(* IEC 61131-3 sources: rusty/libs/stdlib/iec61131-st (part 2) *)

(* ---- num_conversion.st ---- *)
(********************
*
* Converts LREAL to REAL
*
*********************)
FUNCTION LREAL_TO_REAL : REAL
VAR_INPUT
    in : LREAL;
END_VAR
    LREAL_TO_REAL := in;
END_FUNCTION

(********************
*
* Converts LREAL to LINT
*
*********************)
{external}
FUNCTION LREAL_TO_LINT : LINT
VAR_INPUT
    in : LREAL;
END_VAR
END_FUNCTION

(********************
*
* Converts LREAL to DINT
*
*********************)
{external}
FUNCTION LREAL_TO_DINT : DINT
VAR_INPUT
    in : LREAL;
END_VAR
END_FUNCTION

(********************
*
* Converts LREAL to INT
*
*********************)
{external}
FUNCTION LREAL_TO_INT : INT
VAR_INPUT
    in : LREAL;
END_VAR
END_FUNCTION

(********************
*
* Converts LREAL to SINT
*
*********************)
{external}
FUNCTION LREAL_TO_SINT : SINT
VAR_INPUT
    in : LREAL;
END_VAR
END_FUNCTION

(********************
*
* Converts LREAL to ULINT
*
*********************)
{external}
FUNCTION LREAL_TO_ULINT : ULINT
VAR_INPUT
    in : LREAL;
END_VAR
END_FUNCTION

(********************
*
* Converts LREAL to UDINT
*
*********************)
{external}
FUNCTION LREAL_TO_UDINT : UDINT
VAR_INPUT
    in : LREAL;
END_VAR
END_FUNCTION

(********************
*
* Converts LREAL to UINT
*
*********************)
{external}
FUNCTION LREAL_TO_UINT : UINT
VAR_INPUT
    in : LREAL;
END_VAR
END_FUNCTION

(********************
*
* Converts LREAL to USINT
*
*********************)
{external}
FUNCTION LREAL_TO_USINT : USINT
VAR_INPUT
    in : LREAL;
END_VAR
END_FUNCTION

(********************
*
* Converts REAL to LREAL
*
*********************)
FUNCTION REAL_TO_LREAL : LREAL
VAR_INPUT
    in : REAL;
END_VAR
    REAL_TO_LREAL := in;
END_FUNCTION

(********************
*
* Converts REAL to LINT
*
*********************)
{external}
FUNCTION REAL_TO_LINT : LINT
VAR_INPUT
    in : REAL;
END_VAR
END_FUNCTION

(********************
*
* Converts REAL to DINT
*
*********************)
{external}
FUNCTION REAL_TO_DINT : DINT
VAR_INPUT
    in : REAL;
END_VAR
END_FUNCTION

(********************
*
* Converts REAL to INT
*
*********************)
{external}
FUNCTION REAL_TO_INT : INT
VAR_INPUT
    in : REAL;
END_VAR
END_FUNCTION

(********************
*
* Converts REAL to SINT
*
*********************)
{external}
FUNCTION REAL_TO_SINT : SINT
VAR_INPUT
    in : REAL;
END_VAR
END_FUNCTION

(********************
*
* Converts REAL to ULINT
*
*********************)
{external}
FUNCTION REAL_TO_ULINT : ULINT
VAR_INPUT
    in : REAL;
END_VAR
END_FUNCTION

(********************
*
* Converts REAL to UDINT
*
*********************)
{external}
FUNCTION REAL_TO_UDINT : UDINT
VAR_INPUT
    in : REAL;
END_VAR
END_FUNCTION

(********************
*
* Converts REAL to UINT
*
*********************)
{external}
FUNCTION REAL_TO_UINT : UINT
VAR_INPUT
    in : REAL;
END_VAR
END_FUNCTION

(********************
*
* Converts REAL to USINT
*
*********************)
{external}
FUNCTION REAL_TO_USINT : USINT
VAR_INPUT
    in : REAL;
END_VAR
END_FUNCTION

(********************
*
* Converts LINT to LREAL
*
*********************)
FUNCTION LINT_TO_LREAL : LREAL
VAR_INPUT
    in : LINT;
END_VAR
    LINT_TO_LREAL := in;
END_FUNCTION

(********************
*
* Converts LINT to REAL
*
*********************)
FUNCTION LINT_TO_REAL : REAL
VAR_INPUT
    in : LINT;
END_VAR
    LINT_TO_REAL := in;
END_FUNCTION

(********************
*
* Converts LINT to DINT
*
*********************)
FUNCTION LINT_TO_DINT : DINT
VAR_INPUT
    in : LINT;
END_VAR
    LINT_TO_DINT := in;
END_FUNCTION

(********************
*
* Converts LINT to INT
*
*********************)
FUNCTION LINT_TO_INT : INT
VAR_INPUT
    in : LINT;
END_VAR
    LINT_TO_INT := in;
END_FUNCTION

(********************
*
* Converts LINT to SINT
*
*********************)
FUNCTION LINT_TO_SINT : SINT
VAR_INPUT
    in : LINT;
END_VAR
    LINT_TO_SINT := in;
END_FUNCTION

(********************
*
* Converts LINT to ULINT
*
*********************)
FUNCTION LINT_TO_ULINT : ULINT
VAR_INPUT
    in : LINT;
END_VAR
    LINT_TO_ULINT := in;
END_FUNCTION

(********************
*
* Converts LINT to UDINT
*
*********************)
FUNCTION LINT_TO_UDINT : UDINT
VAR_INPUT
    in : LINT;
END_VAR
    LINT_TO_UDINT := in;
END_FUNCTION

(********************
*
* Converts LINT to UINT
*
*********************)
FUNCTION LINT_TO_UINT : UINT
VAR_INPUT
    in : LINT;
END_VAR
    LINT_TO_UINT := in;
END_FUNCTION

(********************
*
* Converts LINT to USINT
*
*********************)
FUNCTION LINT_TO_USINT : USINT
VAR_INPUT
    in : LINT;
END_VAR
    LINT_TO_USINT := in;
END_FUNCTION

(********************
*
* Converts DINT to LREAL
*
*********************)
FUNCTION DINT_TO_LREAL : LREAL
VAR_INPUT
    in : DINT;
END_VAR
    DINT_TO_LREAL := in;
END_FUNCTION

(********************
*
* Converts DINT to REAL
*
*********************)
FUNCTION DINT_TO_REAL : REAL
VAR_INPUT
    in : DINT;
END_VAR
    DINT_TO_REAL := in;
END_FUNCTION

(********************
*
* Converts DINT to LINT
*
*********************)
FUNCTION DINT_TO_LINT : LINT
VAR_INPUT
    in : DINT;
END_VAR
    DINT_TO_LINT := in;
END_FUNCTION

(********************
*
* Converts DINT to INT
*
*********************)
FUNCTION DINT_TO_INT : INT
VAR_INPUT
    in : DINT;
END_VAR
    DINT_TO_INT := in;
END_FUNCTION

(********************
*
* Converts DINT to SINT
*
*********************)
FUNCTION DINT_TO_SINT : SINT
VAR_INPUT
    in : DINT;
END_VAR
    DINT_TO_SINT := in;
END_FUNCTION

(********************
*
* Converts DINT to ULINT
*
*********************)
FUNCTION DINT_TO_ULINT : ULINT
VAR_INPUT
    in : DINT;
END_VAR
    DINT_TO_ULINT := in;
END_FUNCTION

(********************
*
* Converts DINT to UDINT
*
*********************)
FUNCTION DINT_TO_UDINT : UDINT
VAR_INPUT
    in : DINT;
END_VAR
    DINT_TO_UDINT := in;
END_FUNCTION

(********************
*
* Converts DINT to UINT
*
*********************)
FUNCTION DINT_TO_UINT : UINT
VAR_INPUT
    in : DINT;
END_VAR
    DINT_TO_UINT := in;
END_FUNCTION

(********************
*
* Converts DINT to USINT
*
*********************)
FUNCTION DINT_TO_USINT : USINT
VAR_INPUT
    in : DINT;
END_VAR
    DINT_TO_USINT := in;
END_FUNCTION

(********************
*
* Converts INT to LREAL
*
*********************)
FUNCTION INT_TO_LREAL : LREAL
VAR_INPUT
    in : INT;
END_VAR
    INT_TO_LREAL := in;
END_FUNCTION

(********************
*
* Converts INT to REAL
*
*********************)
FUNCTION INT_TO_REAL : REAL
VAR_INPUT
    in : INT;
END_VAR
    INT_TO_REAL := in;
END_FUNCTION

(********************
*
* Converts INT to LINT
*
*********************)
FUNCTION INT_TO_LINT : LINT
VAR_INPUT
    in : INT;
END_VAR
    INT_TO_LINT := in;
END_FUNCTION

(********************
*
* Converts INT to DINT
*
*********************)
FUNCTION INT_TO_DINT : DINT
VAR_INPUT
    in : INT;
END_VAR
    INT_TO_DINT := in;
END_FUNCTION

(********************
*
* Converts INT to SINT
*
*********************)
FUNCTION INT_TO_SINT : SINT
VAR_INPUT
    in : INT;
END_VAR
    INT_TO_SINT := in;
END_FUNCTION

(********************
*
* Converts INT to ULINT
*
*********************)
FUNCTION INT_TO_ULINT : ULINT
VAR_INPUT
    in : INT;
END_VAR
    INT_TO_ULINT := in;
END_FUNCTION

(********************
*
* Converts INT to UDINT
*
*********************)
FUNCTION INT_TO_UDINT : UDINT
VAR_INPUT
    in : INT;
END_VAR
    INT_TO_UDINT := in;
END_FUNCTION

(********************
*
* Converts INT to UINT
*
*********************)
FUNCTION INT_TO_UINT : UINT
VAR_INPUT
    in : INT;
END_VAR
    INT_TO_UINT := in;
END_FUNCTION

(********************
*
* Converts INT to USINT
*
*********************)
FUNCTION INT_TO_USINT : USINT
VAR_INPUT
    in : INT;
END_VAR
    INT_TO_USINT := in;
END_FUNCTION

(********************
*
* Converts SINT to LREAL
*
*********************)
FUNCTION SINT_TO_LREAL : LREAL
VAR_INPUT
    in : SINT;
END_VAR
    SINT_TO_LREAL := in;
END_FUNCTION

(********************
*
* Converts SINT to REAL
*
*********************)
FUNCTION SINT_TO_REAL : REAL
VAR_INPUT
    in : SINT;
END_VAR
    SINT_TO_REAL := in;
END_FUNCTION

(********************
*
* Converts SINT to LINT
*
*********************)
FUNCTION SINT_TO_LINT : LINT
VAR_INPUT
    in : SINT;
END_VAR
    SINT_TO_LINT := in;
END_FUNCTION

(********************
*
* Converts SINT to DINT
*
*********************)
FUNCTION SINT_TO_DINT : DINT
VAR_INPUT
    in : SINT;
END_VAR
    SINT_TO_DINT := in;
END_FUNCTION

(********************
*
* Converts SINT to INT
*
*********************)
FUNCTION SINT_TO_INT : INT
VAR_INPUT
    in : SINT;
END_VAR
    SINT_TO_INT := in;
END_FUNCTION

(********************
*
* Converts SINT to ULINT
*
*********************)
FUNCTION SINT_TO_ULINT : ULINT
VAR_INPUT
    in : SINT;
END_VAR
    SINT_TO_ULINT := in;
END_FUNCTION

(********************
*
* Converts SINT to UDINT
*
*********************)
FUNCTION SINT_TO_UDINT : UDINT
VAR_INPUT
    in : SINT;
END_VAR
    SINT_TO_UDINT := in;
END_FUNCTION

(********************
*
* Converts SINT to UINT
*
*********************)
FUNCTION SINT_TO_UINT : UINT
VAR_INPUT
    in : SINT;
END_VAR
    SINT_TO_UINT := in;
END_FUNCTION

(********************
*
* Converts SINT to USINT
*
*********************)
FUNCTION SINT_TO_USINT : USINT
VAR_INPUT
    in : SINT;
END_VAR
    SINT_TO_USINT := in;
END_FUNCTION

(********************
*
* Converts ULINT to LREAL
*
*********************)
FUNCTION ULINT_TO_LREAL : LREAL
VAR_INPUT
    in : ULINT;
END_VAR
    ULINT_TO_LREAL := in;
END_FUNCTION

(********************
*
* Converts ULINT to REAL
*
*********************)
FUNCTION ULINT_TO_REAL : REAL
VAR_INPUT
    in : ULINT;
END_VAR
    ULINT_TO_REAL := in;
END_FUNCTION

(********************
*
* Converts ULINT to LINT
*
*********************)
FUNCTION ULINT_TO_LINT : LINT
VAR_INPUT
    in : ULINT;
END_VAR
    ULINT_TO_LINT := in;
END_FUNCTION

(********************
*
* Converts ULINT to DINT
*
*********************)
FUNCTION ULINT_TO_DINT : DINT
VAR_INPUT
    in : ULINT;
END_VAR
    ULINT_TO_DINT := in;
END_FUNCTION

(********************
*
* Converts ULINT to INT
*
*********************)
FUNCTION ULINT_TO_INT : INT
VAR_INPUT
    in : ULINT;
END_VAR
    ULINT_TO_INT := in;
END_FUNCTION

(********************
*
* Converts ULINT to SINT
*
*********************)
FUNCTION ULINT_TO_SINT : SINT
VAR_INPUT
    in : ULINT;
END_VAR
    ULINT_TO_SINT := in;
END_FUNCTION

(********************
*
* Converts ULINT to UDINT
*
*********************)
FUNCTION ULINT_TO_UDINT : UDINT
VAR_INPUT
    in : ULINT;
END_VAR
    ULINT_TO_UDINT := in;
END_FUNCTION

(********************
*
* Converts ULINT to UINT
*
*********************)
FUNCTION ULINT_TO_UINT : UINT
VAR_INPUT
    in : ULINT;
END_VAR
    ULINT_TO_UINT := in;
END_FUNCTION

(********************
*
* Converts ULINT to USINT
*
*********************)
FUNCTION ULINT_TO_USINT : USINT
VAR_INPUT
    in : ULINT;
END_VAR
    ULINT_TO_USINT := in;
END_FUNCTION

(********************
*
* Converts UDINT to LREAL
*
*********************)
FUNCTION UDINT_TO_LREAL : LREAL
VAR_INPUT
    in : UDINT;
END_VAR
    UDINT_TO_LREAL := in;
END_FUNCTION

(********************
*
* Converts UDINT to REAL
*
*********************)
FUNCTION UDINT_TO_REAL : REAL
VAR_INPUT
    in : UDINT;
END_VAR
    UDINT_TO_REAL := in;
END_FUNCTION

(********************
*
* Converts UDINT to LINT
*
*********************)
FUNCTION UDINT_TO_LINT : LINT
VAR_INPUT
    in : UDINT;
END_VAR
    UDINT_TO_LINT := in;
END_FUNCTION

(********************
*
* Converts UDINT to DINT
*
*********************)
FUNCTION UDINT_TO_DINT : DINT
VAR_INPUT
    in : UDINT;
END_VAR
    UDINT_TO_DINT := in;
END_FUNCTION

(********************
*
* Converts UDINT to INT
*
*********************)
FUNCTION UDINT_TO_INT : INT
VAR_INPUT
    in : UDINT;
END_VAR
    UDINT_TO_INT := in;
END_FUNCTION

(********************
*
* Converts UDINT to SINT
*
*********************)
FUNCTION UDINT_TO_SINT : SINT
VAR_INPUT
    in : UDINT;
END_VAR
    UDINT_TO_SINT := in;
END_FUNCTION

(********************
*
* Converts UDINT to ULINT
*
*********************)
FUNCTION UDINT_TO_ULINT : ULINT
VAR_INPUT
    in : UDINT;
END_VAR
    UDINT_TO_ULINT := in;
END_FUNCTION

(********************
*
* Converts UDINT to UINT
*
*********************)
FUNCTION UDINT_TO_UINT : UINT
VAR_INPUT
    in : UDINT;
END_VAR
    UDINT_TO_UINT := in;
END_FUNCTION

(********************
*
* Converts UDINT to USINT
*
*********************)
FUNCTION UDINT_TO_USINT : USINT
VAR_INPUT
    in : UDINT;
END_VAR
    UDINT_TO_USINT := in;
END_FUNCTION

(********************
*
* Converts UINT to LREAL
*
*********************)
FUNCTION UINT_TO_LREAL : LREAL
VAR_INPUT
    in : UINT;
END_VAR
    UINT_TO_LREAL := in;
END_FUNCTION

(********************
*
* Converts UINT to REAL
*
*********************)
FUNCTION UINT_TO_REAL : REAL
VAR_INPUT
    in : UINT;
END_VAR
    UINT_TO_REAL := in;
END_FUNCTION

(********************
*
* Converts UINT to LINT
*
*********************)
FUNCTION UINT_TO_LINT : LINT
VAR_INPUT
    in : UINT;
END_VAR
    UINT_TO_LINT := in;
END_FUNCTION

(********************
*
* Converts UINT to DINT
*
*********************)
FUNCTION UINT_TO_DINT : DINT
VAR_INPUT
    in : UINT;
END_VAR
    UINT_TO_DINT := in;
END_FUNCTION

(********************
*
* Converts UINT to INT
*
*********************)
FUNCTION UINT_TO_INT : INT
VAR_INPUT
    in : UINT;
END_VAR
    UINT_TO_INT := in;
END_FUNCTION

(********************
*
* Converts UINT to SINT
*
*********************)
FUNCTION UINT_TO_SINT : SINT
VAR_INPUT
    in : UINT;
END_VAR
    UINT_TO_SINT := in;
END_FUNCTION

(********************
*
* Converts UINT to ULINT
*
*********************)
FUNCTION UINT_TO_ULINT : ULINT
VAR_INPUT
    in : UINT;
END_VAR
    UINT_TO_ULINT := in;
END_FUNCTION

(********************
*
* Converts UINT to UDINT
*
*********************)
FUNCTION UINT_TO_UDINT : UDINT
VAR_INPUT
    in : UINT;
END_VAR
    UINT_TO_UDINT := in;
END_FUNCTION

(********************
*
* Converts UINT to USINT
*
*********************)
FUNCTION UINT_TO_USINT : USINT
VAR_INPUT
    in : UINT;
END_VAR
    UINT_TO_USINT := in;
END_FUNCTION

(********************
*
* Converts USINT to LREAL
*
*********************)
FUNCTION USINT_TO_LREAL : LREAL
VAR_INPUT
    in : USINT;
END_VAR
    USINT_TO_LREAL := in;
END_FUNCTION

(********************
*
* Converts USINT to REAL
*
*********************)
FUNCTION USINT_TO_REAL : REAL
VAR_INPUT
    in : USINT;
END_VAR
    USINT_TO_REAL := in;
END_FUNCTION

(********************
*
* Converts USINT to LINT
*
*********************)
FUNCTION USINT_TO_LINT : LINT
VAR_INPUT
    in : USINT;
END_VAR
    USINT_TO_LINT := in;
END_FUNCTION

(********************
*
* Converts USINT to DINT
*
*********************)
FUNCTION USINT_TO_DINT : DINT
VAR_INPUT
    in : USINT;
END_VAR
    USINT_TO_DINT := in;
END_FUNCTION

(********************
*
* Converts USINT to INT
*
*********************)
FUNCTION USINT_TO_INT : INT
VAR_INPUT
    in : USINT;
END_VAR
    USINT_TO_INT := in;
END_FUNCTION

(********************
*
* Converts USINT to SINT
*
*********************)
FUNCTION USINT_TO_SINT : SINT
VAR_INPUT
    in : USINT;
END_VAR
    USINT_TO_SINT := in;
END_FUNCTION

(********************
*
* Converts USINT to ULINT
*
*********************)
FUNCTION USINT_TO_ULINT : ULINT
VAR_INPUT
    in : USINT;
END_VAR
    USINT_TO_ULINT := in;
END_FUNCTION

(********************
*
* Converts USINT to UDINT
*
*********************)
FUNCTION USINT_TO_UDINT : UDINT
VAR_INPUT
    in : USINT;
END_VAR
    USINT_TO_UDINT := in;
END_FUNCTION

(********************
*
* Converts USINT to UINT
*
*********************)
FUNCTION USINT_TO_UINT : UINT
VAR_INPUT
    in : USINT;
END_VAR
    USINT_TO_UINT := in;
END_FUNCTION

(* ---- numerical_functions.st ---- *)
(**************************
 *
 *This operator returns the absolute value of a number.
 *
*************************)
FUNCTION ABS<T : ANY_NUM> : T
VAR_INPUT
    IN : T;
END_VAR

END_FUNCTION

(* Specialized implementation of ABS for DINT *)
/* FUNCTION ABS__DINT : DINT */
FUNCTION ABS__DINT : DINT
VAR_INPUT
    IN : DINT;
END_VAR
    ABS__DINT := IN;
    IF ABS__DINT < 0 THEN
        ABS__DINT := -1 * ABS__DINT;
    END_IF
END_FUNCTION

(* Specialized implementation of ABS for SINT *)
FUNCTION ABS__SINT : SINT
VAR_INPUT
    IN : SINT;
END_VAR
    ABS__SINT := ABS__DINT(IN);
END_FUNCTION

(* Specialized implementation of ABS for INT *)
FUNCTION ABS__INT : INT
VAR_INPUT
    IN : INT;
END_VAR
    ABS__INT := ABS__DINT(IN);
END_FUNCTION

(* Specialized implementation of ABS for LINT *)
FUNCTION ABS__LINT : LINT
VAR_INPUT
    IN : LINT;
END_VAR
    ABS__LINT := IN;
    IF ABS__LINT < 0 THEN
        ABS__LINT := -1 * ABS__LINT;
    END_IF
END_FUNCTION

(* Specialized implementation of ABS for REAL *)
FUNCTION ABS__REAL : REAL
VAR_INPUT
    IN : REAL;
END_VAR
    ABS__REAL := ABS__LREAL(IN);
END_FUNCTION

(* Specialized implementation of ABS for LREAL *)
FUNCTION ABS__LREAL : LREAL
VAR_INPUT
    IN : LREAL;
END_VAR
    ABS__LREAL := IN;
    IF ABS__LREAL < 0 THEN
        ABS__LREAL := -1.0 * ABS__LREAL;
    END_IF
END_FUNCTION

(* ---- real_trunc_int.st ---- *)
(********************
*
* Converts REAL to SINT
*
********************)
FUNCTION REAL_TRUNC_SINT : SINT
    VAR_INPUT
        in : REAL;
    END_VAR

    REAL_TRUNC_SINT := in;
END_FUNCTION

(********************
*
* Converts REAL to USINT
*
********************)
FUNCTION REAL_TRUNC_USINT : USINT
    VAR_INPUT
        in : REAL;
    END_VAR

    REAL_TRUNC_USINT := in;
END_FUNCTION

(********************
*
* Converts REAL to INT
*
********************)
FUNCTION REAL_TRUNC_INT : INT
    VAR_INPUT
        in : REAL;
    END_VAR

    REAL_TRUNC_INT := in;
END_FUNCTION

(********************
*
* Converts REAL to UINT
*
********************)
FUNCTION REAL_TRUNC_UINT : UINT
    VAR_INPUT
        in : REAL;
    END_VAR

    REAL_TRUNC_UINT := in;
END_FUNCTION

(********************
*
* Converts REAL to DINT
*
********************)
FUNCTION REAL_TRUNC_DINT : DINT
    VAR_INPUT
        in : REAL;
    END_VAR

    REAL_TRUNC_DINT := in;
END_FUNCTION

(********************
*
* Converts REAL to UDINT
*
********************)
FUNCTION REAL_TRUNC_UDINT : UDINT
    VAR_INPUT
        in : REAL;
    END_VAR

    REAL_TRUNC_UDINT := in;
END_FUNCTION

(********************
*
* Converts REAL to LINT
*
********************)
FUNCTION REAL_TRUNC_LINT : LINT
    VAR_INPUT
        in : REAL;
    END_VAR

    REAL_TRUNC_LINT := in;
END_FUNCTION

(********************
*
* Converts REAL to ULINT
*
********************)
FUNCTION REAL_TRUNC_ULINT : ULINT
    VAR_INPUT
        in : REAL;
    END_VAR

    REAL_TRUNC_ULINT := in;
END_FUNCTION

(********************
*
* Converts LREAL to SINT
*
********************)
FUNCTION LREAL_TRUNC_SINT : SINT
    VAR_INPUT
        in : LREAL;
    END_VAR

    LREAL_TRUNC_SINT := in;
END_FUNCTION

(********************
*
* Converts LREAL to USINT
*
********************)
FUNCTION LREAL_TRUNC_USINT : USINT
    VAR_INPUT
        in : LREAL;
    END_VAR

    LREAL_TRUNC_USINT := in;
END_FUNCTION

(********************
*
* Converts LREAL to INT
*
********************)
FUNCTION LREAL_TRUNC_INT : INT
    VAR_INPUT
        in : LREAL;
    END_VAR

    LREAL_TRUNC_INT := in;
END_FUNCTION

(********************
*
* Converts LREAL to UINT
*
********************)
FUNCTION LREAL_TRUNC_UINT : UINT
    VAR_INPUT
        in : LREAL;
    END_VAR

    LREAL_TRUNC_UINT := in;
END_FUNCTION

(********************
*
* Converts LREAL to DINT
*
********************)
FUNCTION LREAL_TRUNC_DINT : DINT
    VAR_INPUT
        in : LREAL;
    END_VAR

    LREAL_TRUNC_DINT := in;
END_FUNCTION

(********************
*
* Converts LREAL to UDINT
*
********************)
FUNCTION LREAL_TRUNC_UDINT : UDINT
    VAR_INPUT
        in : LREAL;
    END_VAR

    LREAL_TRUNC_UDINT := in;
END_FUNCTION

(********************
*
* Converts LREAL to LINT
*
********************)
FUNCTION LREAL_TRUNC_LINT : LINT
    VAR_INPUT
        in : LREAL;
    END_VAR

    LREAL_TRUNC_LINT := in;
END_FUNCTION

(********************
*
* Converts LREAL to ULINT
*
********************)
FUNCTION LREAL_TRUNC_ULINT : ULINT
    VAR_INPUT
        in : LREAL;
    END_VAR

    LREAL_TRUNC_ULINT := in;
END_FUNCTION

(* ---- selectors.st ---- *)
(**************************
 *
 * MAX(IN0, IN1, ...)
 *
 * This operator produces the larger value of the given operands.
 *
*************************)
{external}
FUNCTION MAX<T: ANY_ELEMENTARY> : T
VAR_INPUT
    IN : {sized} T...;
END_VAR
END_FUNCTION

(**************************
 *
 * MIN(IN0, IN1, ...)
 *
 * This operator produces the smaller value of the given operands.
 *
*************************)
{external}
FUNCTION MIN<T: ANY_ELEMENTARY> : T
VAR_INPUT
    IN : {sized} T...;
END_VAR
END_FUNCTION

(**************************
 *
 * LIMIT(Min, IN, Max)
 *
 * This operator limits an input value to the range between Min and Max.
 * If IN lies between the range of Min and Max, IN is displayed as a result.
 * If IN > Max, Max is displayed as a result.
 * If IN < Min, Min is displayed as a result.
 *
*************************)
{external}
FUNCTION LIMIT<T: ANY_ELEMENTARY> : T
VAR_INPUT
    MIN : T;
    IN : T;
    MAX : T;
END_VAR
END_FUNCTION

(* ---- string_conversion.st ---- *)
(********************
*
* Converts WSTRING to STRING
*
*********************)
FUNCTION WSTRING_TO_STRING : STRING[__STRING_LENGTH]
VAR_INPUT {ref}
    in : WSTRING[__STRING_LENGTH];
END_VAR
    WSTRING_TO_STRING_EXT(in, WSTRING_TO_STRING);
END_FUNCTION

{external}
FUNCTION WSTRING_TO_STRING_EXT : DINT
VAR_INPUT {ref}
    in : WSTRING[__STRING_LENGTH];
END_VAR
VAR_IN_OUT
    out : STRING[__STRING_LENGTH];
END_VAR
END_FUNCTION

(********************
*
* Converts WSTRING to WCHAR
*
*********************)
{external}
FUNCTION WSTRING_TO_WCHAR : WCHAR
VAR_INPUT {ref}
    in : WSTRING;
END_VAR
END_FUNCTION

(********************
*
* Converts STRING to WSTRING
* Will return a WSTRING with default length of 81
*
*********************)
FUNCTION STRING_TO_WSTRING : WSTRING[__STRING_LENGTH]
VAR_INPUT {ref}
    in : STRING[__STRING_LENGTH];
END_VAR
    STRING_TO_WSTRING_EXT(in, STRING_TO_WSTRING);
END_FUNCTION

{external}
FUNCTION STRING_TO_WSTRING_EXT : DINT
VAR_INPUT {ref}
    in : STRING[__STRING_LENGTH];
END_VAR
VAR_IN_OUT
    out : WSTRING[__STRING_LENGTH];
END_VAR
END_FUNCTION

(********************
*
* Converts STRING to CHAR
*
*********************)
{external}
FUNCTION STRING_TO_CHAR : CHAR
VAR_INPUT {ref}
    in : STRING;
END_VAR
END_FUNCTION

(********************
*
* Converts WCHAR to WSTRING
*
*********************)
{external}
FUNCTION WCHAR_TO_WSTRING : WSTRING
VAR_INPUT
    in : WCHAR;
END_VAR
END_FUNCTION

(********************
*
* Converts WCHAR to CHAR
*
*********************)
{external}
FUNCTION WCHAR_TO_CHAR : CHAR
VAR_INPUT
    in : WCHAR;
END_VAR
END_FUNCTION

(********************
*
* Converts CHAR to STRING
*
*********************)
{external}
FUNCTION CHAR_TO_STRING : STRING
VAR_INPUT
    in : CHAR;
END_VAR
END_FUNCTION

(********************
*
* Converts CHAR to WCHAR
*
*********************)
{external}
FUNCTION CHAR_TO_WCHAR : WCHAR
VAR_INPUT
    in : CHAR;
END_VAR
END_FUNCTION

(* ---- string_to_conversions.st ---- *)
(******************************************************************************
*
* Converts STRING and WSTRING values to native values.
*
******************************************************************************)

(******************************************************************************
*
* Converts STRING to BOOL. Never faults; a rejected input yields FALSE.
*
******************************************************************************)
{external}
FUNCTION STRING_TO_BOOL : BOOL
VAR_INPUT {ref}
    IN : STRING;
END_VAR
END_FUNCTION

(******************************************************************************
*
* Converts STRING to BYTE. Never faults; a rejected input yields 0.
*
******************************************************************************)
{external}
FUNCTION STRING_TO_BYTE : BYTE
VAR_INPUT {ref}
    IN : STRING;
END_VAR
END_FUNCTION

(******************************************************************************
*
* Converts STRING to WORD. Never faults; a rejected input yields 0.
*
******************************************************************************)
{external}
FUNCTION STRING_TO_WORD : WORD
VAR_INPUT {ref}
    IN : STRING;
END_VAR
END_FUNCTION

(******************************************************************************
*
* Converts STRING to DWORD. Never faults; a rejected input yields 0.
*
******************************************************************************)
{external}
FUNCTION STRING_TO_DWORD : DWORD
VAR_INPUT {ref}
    IN : STRING;
END_VAR
END_FUNCTION

(******************************************************************************
*
* Converts STRING to LWORD. Never faults; a rejected input yields 0.
*
******************************************************************************)
{external}
FUNCTION STRING_TO_LWORD : LWORD
VAR_INPUT {ref}
    IN : STRING;
END_VAR
END_FUNCTION

(******************************************************************************
*
* Converts STRING to SINT. Never faults; a rejected input yields 0.
*
******************************************************************************)
{external}
FUNCTION STRING_TO_SINT : SINT
VAR_INPUT {ref}
    IN : STRING;
END_VAR
END_FUNCTION

(******************************************************************************
*
* Converts STRING to USINT. Never faults; a rejected input yields 0.
*
******************************************************************************)
{external}
FUNCTION STRING_TO_USINT : USINT
VAR_INPUT {ref}
    IN : STRING;
END_VAR
END_FUNCTION

(******************************************************************************
*
* Converts STRING to INT. Never faults; a rejected input yields 0.
*
******************************************************************************)
{external}
FUNCTION STRING_TO_INT : INT
VAR_INPUT {ref}
    IN : STRING;
END_VAR
END_FUNCTION

(******************************************************************************
*
* Converts STRING to UINT. Never faults; a rejected input yields 0.
*
******************************************************************************)
{external}
FUNCTION STRING_TO_UINT : UINT
VAR_INPUT {ref}
    IN : STRING;
END_VAR
END_FUNCTION

(******************************************************************************
*
* Converts STRING to DINT. Never faults; a rejected input yields 0.
*
******************************************************************************)
{external}
FUNCTION STRING_TO_DINT : DINT
VAR_INPUT {ref}
    IN : STRING;
END_VAR
END_FUNCTION

(******************************************************************************
*
* Converts STRING to UDINT. Never faults; a rejected input yields 0.
*
******************************************************************************)
{external}
FUNCTION STRING_TO_UDINT : UDINT
VAR_INPUT {ref}
    IN : STRING;
END_VAR
END_FUNCTION

(******************************************************************************
*
* Converts STRING to LINT. Never faults; a rejected input yields 0.
*
******************************************************************************)
{external}
FUNCTION STRING_TO_LINT : LINT
VAR_INPUT {ref}
    IN : STRING;
END_VAR
END_FUNCTION

(******************************************************************************
*
* Converts STRING to ULINT. Never faults; a rejected input yields 0.
*
******************************************************************************)
{external}
FUNCTION STRING_TO_ULINT : ULINT
VAR_INPUT {ref}
    IN : STRING;
END_VAR
END_FUNCTION

(******************************************************************************
*
* Converts STRING to LREAL.
*
******************************************************************************)
{external}
FUNCTION STRING_TO_LREAL : LREAL
VAR_INPUT {ref}
    IN : STRING;
END_VAR
END_FUNCTION

(******************************************************************************
*
* Converts STRING to REAL.
*
******************************************************************************)
{external}
FUNCTION STRING_TO_REAL : REAL
VAR_INPUT {ref}
    IN : STRING;
END_VAR
END_FUNCTION

(******************************************************************************
*
* Converts STRING to TIME. Requires a T#/TIME# prefix; never faults, a rejected or
* negative duration yields T#0s.
*
******************************************************************************)
{external}
FUNCTION STRING_TO_TIME : TIME
VAR_INPUT {ref}
    IN : STRING;
END_VAR
END_FUNCTION

(******************************************************************************
*
* Converts STRING to LTIME. Requires a LT#/LTIME# prefix; never faults, a rejected or
* negative duration yields LTIME#0s.
*
******************************************************************************)
{external}
FUNCTION STRING_TO_LTIME : LTIME
VAR_INPUT {ref}
    IN : STRING;
END_VAR
END_FUNCTION

(******************************************************************************
*
* Converts STRING to DATE. Requires a D#/DATE# prefix. Never faults; an impossible or
* out-of-range (1970-01-01..2106-02-07) date yields D#1970-01-01.
*
******************************************************************************)
{external}
FUNCTION STRING_TO_DATE : DATE
VAR_INPUT {ref}
    IN : STRING;
END_VAR
END_FUNCTION

(******************************************************************************
*
* Converts STRING to DT. Requires a DT#/DATE_AND_TIME# prefix. Never faults; an
* impossible or out-of-range date-time yields DT#1970-01-01-00:00:00.
*
******************************************************************************)
{external}
FUNCTION STRING_TO_DT : DT
VAR_INPUT {ref}
    IN : STRING;
END_VAR
END_FUNCTION

(******************************************************************************
*
* Converts STRING to TOD. Requires a TOD#/TIME_OF_DAY# prefix. Never faults; an
* impossible time yields TOD#00:00:00.
*
******************************************************************************)
{external}
FUNCTION STRING_TO_TOD : TOD
VAR_INPUT {ref}
    IN : STRING;
END_VAR
END_FUNCTION

(******************************************************************************
*
* Converts WSTRING to LINT.
*
******************************************************************************)
FUNCTION WSTRING_TO_LINT : LINT
VAR_INPUT {ref}
    IN : WSTRING;
END_VAR
VAR_TEMP
    STR : STRING;
END_VAR
    WSTRING_TO_STRING_EXT(IN, STR);
    WSTRING_TO_LINT := STRING_TO_LINT(STR);
END_FUNCTION

(******************************************************************************
*
* Converts WSTRING to DINT.
*
******************************************************************************)
FUNCTION WSTRING_TO_DINT : DINT
VAR_INPUT {ref}
    IN : WSTRING;
END_VAR
VAR_TEMP
    STR : STRING;
END_VAR
    WSTRING_TO_STRING_EXT(IN, STR);
    WSTRING_TO_DINT := STRING_TO_DINT(STR);
END_FUNCTION

(******************************************************************************
*
* Converts WSTRING to LREAL.
*
******************************************************************************)
FUNCTION WSTRING_TO_LREAL : LREAL
VAR_INPUT {ref}
    IN : WSTRING;
END_VAR
VAR_TEMP
    STR : STRING;
END_VAR
    WSTRING_TO_STRING_EXT(IN, STR);
    WSTRING_TO_LREAL := STRING_TO_LREAL(STR);
END_FUNCTION

(******************************************************************************
*
* Converts WSTRING to REAL.
*
******************************************************************************)
FUNCTION WSTRING_TO_REAL : REAL
VAR_INPUT {ref}
    IN : WSTRING;
END_VAR
VAR_TEMP
    STR : STRING;
END_VAR
    WSTRING_TO_STRING_EXT(IN, STR);
    WSTRING_TO_REAL := STRING_TO_REAL(STR);
END_FUNCTION

(* ---- to_bit.st ---- *)
FUNCTION TO_BOOL<T: ANY> : BOOL
    VAR_INPUT
        in : T;
    END_VAR
END_FUNCTION

FUNCTION TO_BOOL__BOOL : BOOL
    VAR_INPUT
        in : BOOL;
    END_VAR

    TO_BOOL__BOOL := in;
END_FUNCTION

FUNCTION TO_BOOL__BYTE : BOOL
    VAR_INPUT
        in : BYTE;
    END_VAR

    TO_BOOL__BYTE := BYTE_TO_BOOL(in);
END_FUNCTION

FUNCTION TO_BOOL__WORD : BOOL
    VAR_INPUT
        in : WORD;
    END_VAR

    TO_BOOL__WORD := WORD_TO_BOOL(in);
END_FUNCTION

FUNCTION TO_BOOL__DWORD : BOOL
    VAR_INPUT
        in : DWORD;
    END_VAR

    TO_BOOL__DWORD := DWORD_TO_BOOL(in);
END_FUNCTION

FUNCTION TO_BOOL__LWORD : BOOL
    VAR_INPUT
        in : LWORD;
    END_VAR

    TO_BOOL__LWORD := LWORD_TO_BOOL(in);
END_FUNCTION

FUNCTION TO_BOOL__SINT : BOOL
    VAR_INPUT
        in : SINT;
    END_VAR

    TO_BOOL__SINT := SINT_TO_BOOL(in);
END_FUNCTION

FUNCTION TO_BOOL__USINT : BOOL
    VAR_INPUT
        in : USINT;
    END_VAR

    TO_BOOL__USINT := USINT_TO_BOOL(in);
END_FUNCTION

FUNCTION TO_BOOL__INT : BOOL
    VAR_INPUT
        in : INT;
    END_VAR

    TO_BOOL__INT := INT_TO_BOOL(in);
END_FUNCTION

FUNCTION TO_BOOL__UINT : BOOL
    VAR_INPUT
        in : UINT;
    END_VAR

    TO_BOOL__UINT := UINT_TO_BOOL(in);
END_FUNCTION

FUNCTION TO_BOOL__DINT : BOOL
    VAR_INPUT
        in : DINT;
    END_VAR

    TO_BOOL__DINT := DINT_TO_BOOL(in);
END_FUNCTION

FUNCTION TO_BOOL__UDINT : BOOL
    VAR_INPUT
        in : UDINT;
    END_VAR

    TO_BOOL__UDINT := UDINT_TO_BOOL(in);
END_FUNCTION

FUNCTION TO_BOOL__LINT : BOOL
    VAR_INPUT
        in : LINT;
    END_VAR

    TO_BOOL__LINT := LINT_TO_BOOL(in);
END_FUNCTION

FUNCTION TO_BOOL__ULINT : BOOL
    VAR_INPUT
        in : ULINT;
    END_VAR

    TO_BOOL__ULINT := ULINT_TO_BOOL(in);
END_FUNCTION

FUNCTION TO_BOOL__REAL : BOOL
    VAR_INPUT
        in : REAL;
    END_VAR

    TO_BOOL__REAL := REAL_TO_BOOL(in);
END_FUNCTION

FUNCTION TO_BOOL__LREAL : BOOL
    VAR_INPUT
        in : LREAL;
    END_VAR

    TO_BOOL__LREAL := LREAL_TO_BOOL(in);
END_FUNCTION

// ======================================================================================================== //

FUNCTION TO_BYTE<T: ANY> : BYTE
    VAR_INPUT
        in : T;
    END_VAR
END_FUNCTION

FUNCTION TO_BYTE__BYTE : BYTE
    VAR_INPUT
        in : BYTE;
    END_VAR

    TO_BYTE__BYTE := in;
END_FUNCTION

FUNCTION TO_BYTE__BOOL : BYTE
    VAR_INPUT
        in : BOOL;
    END_VAR

    TO_BYTE__BOOL := BOOL_TO_BYTE(in);
END_FUNCTION

FUNCTION TO_BYTE__CHAR : BYTE
    VAR_INPUT
        in : CHAR;
    END_VAR

    TO_BYTE__CHAR := CHAR_TO_BYTE(in);
END_FUNCTION

FUNCTION TO_BYTE__WCHAR : BYTE
    VAR_INPUT
        in : WCHAR;
    END_VAR

    TO_BYTE__WCHAR := WCHAR_TO_BYTE(in);
END_FUNCTION

FUNCTION TO_BYTE__WORD : BYTE
    VAR_INPUT
        in : WORD;
    END_VAR

    TO_BYTE__WORD := WORD_TO_BYTE(in);
END_FUNCTION

FUNCTION TO_BYTE__DWORD : BYTE
    VAR_INPUT
        in : DWORD;
    END_VAR

    TO_BYTE__DWORD := DWORD_TO_BYTE(in);
END_FUNCTION

FUNCTION TO_BYTE__LWORD : BYTE
    VAR_INPUT
        in : LWORD;
    END_VAR

    TO_BYTE__LWORD := LWORD_TO_BYTE(in);
END_FUNCTION

FUNCTION TO_BYTE__REAL : BYTE
    VAR_INPUT
        in : REAL;
    END_VAR

    TO_BYTE__REAL := REAL_TO_BYTE(in);
END_FUNCTION

FUNCTION TO_BYTE__LREAL : BYTE
    VAR_INPUT
        in : LREAL;
    END_VAR

    TO_BYTE__LREAL := LREAL_TO_BYTE(in);
END_FUNCTION

// ======================================================================================================== //

FUNCTION TO_WORD<T: ANY> : WORD
    VAR_INPUT
        in : T;
    END_VAR
END_FUNCTION

FUNCTION TO_WORD__WORD : WORD
    VAR_INPUT
        in : WORD;
    END_VAR

    TO_WORD__WORD := in;
END_FUNCTION

FUNCTION TO_WORD__BOOL : WORD
    VAR_INPUT
        in : BOOL;
    END_VAR

    TO_WORD__BOOL := BOOL_TO_WORD(in);
END_FUNCTION

FUNCTION TO_WORD__CHAR : WORD
    VAR_INPUT
        in : CHAR;
    END_VAR

    TO_WORD__CHAR := CHAR_TO_WORD(in);
END_FUNCTION

FUNCTION TO_WORD__WCHAR : WORD
    VAR_INPUT
        in : WCHAR;
    END_VAR

    TO_WORD__WCHAR := WCHAR_TO_WORD(in);
END_FUNCTION

FUNCTION TO_WORD__BYTE : WORD
    VAR_INPUT
        in : BYTE;
    END_VAR

    TO_WORD__BYTE := BYTE_TO_WORD(in);
END_FUNCTION

FUNCTION TO_WORD__DWORD : WORD
    VAR_INPUT
        in : DWORD;
    END_VAR

    TO_WORD__DWORD := DWORD_TO_WORD(in);
END_FUNCTION

FUNCTION TO_WORD__LWORD : WORD
    VAR_INPUT
        in : LWORD;
    END_VAR

    TO_WORD__LWORD := LWORD_TO_WORD(in);
END_FUNCTION

FUNCTION TO_WORD__REAL : WORD
    VAR_INPUT
        in : REAL;
    END_VAR

    TO_WORD__REAL := REAL_TO_WORD(in);
END_FUNCTION

FUNCTION TO_WORD__LREAL : WORD
    VAR_INPUT
        in : LREAL;
    END_VAR

    TO_WORD__LREAL := LREAL_TO_WORD(in);
END_FUNCTION

// ======================================================================================================== //

FUNCTION TO_DWORD<T: ANY> : DWORD
    VAR_INPUT
        in : T;
    END_VAR
END_FUNCTION

FUNCTION TO_DWORD__DWORD : DWORD
    VAR_INPUT
        in : DWORD;
    END_VAR

    TO_DWORD__DWORD := in;
END_FUNCTION

FUNCTION TO_DWORD__BOOL : DWORD
    VAR_INPUT
        in : BOOL;
    END_VAR

    TO_DWORD__BOOL := BOOL_TO_DWORD(in);
END_FUNCTION

FUNCTION TO_DWORD__CHAR : DWORD
    VAR_INPUT
        in : CHAR;
    END_VAR

    TO_DWORD__CHAR := CHAR_TO_DWORD(in);
END_FUNCTION

FUNCTION TO_DWORD__WCHAR : DWORD
    VAR_INPUT
        in : WCHAR;
    END_VAR

    TO_DWORD__WCHAR := WCHAR_TO_DWORD(in);
END_FUNCTION

FUNCTION TO_DWORD__BYTE : DWORD
    VAR_INPUT
        in : BYTE;
    END_VAR

    TO_DWORD__BYTE := BYTE_TO_DWORD(in);
END_FUNCTION

FUNCTION TO_DWORD__WORD : DWORD
    VAR_INPUT
        in : WORD;
    END_VAR

    TO_DWORD__WORD := WORD_TO_DWORD(in);
END_FUNCTION

FUNCTION TO_DWORD__LWORD : DWORD
    VAR_INPUT
        in : LWORD;
    END_VAR

    TO_DWORD__LWORD := LWORD_TO_DWORD(in);
END_FUNCTION

FUNCTION TO_DWORD__REAL : DWORD
    VAR_INPUT
        in : REAL;
    END_VAR

    TO_DWORD__REAL := REAL_TO_DWORD(in);
END_FUNCTION

FUNCTION TO_DWORD__LREAL : DWORD
    VAR_INPUT
        in : LREAL;
    END_VAR

    TO_DWORD__LREAL := LREAL_TO_DWORD(in);
END_FUNCTION

// ======================================================================================================== //

FUNCTION TO_LWORD<T: ANY> : LWORD
    VAR_INPUT
        in : T;
    END_VAR
END_FUNCTION

FUNCTION TO_LWORD__LWORD : LWORD
    VAR_INPUT
        in : LWORD;
    END_VAR

    TO_LWORD__LWORD := in;
END_FUNCTION

FUNCTION TO_LWORD__BOOL : LWORD
    VAR_INPUT
        in : BOOL;
    END_VAR

    TO_LWORD__BOOL := BOOL_TO_LWORD(in);
END_FUNCTION

FUNCTION TO_LWORD__CHAR : LWORD
    VAR_INPUT
        in : CHAR;
    END_VAR

    TO_LWORD__CHAR := CHAR_TO_LWORD(in);
END_FUNCTION

FUNCTION TO_LWORD__WCHAR : LWORD
    VAR_INPUT
        in : WCHAR;
    END_VAR

    TO_LWORD__WCHAR := WCHAR_TO_LWORD(in);
END_FUNCTION

FUNCTION TO_LWORD__BYTE : LWORD
    VAR_INPUT
        in : BYTE;
    END_VAR

    TO_LWORD__BYTE := BYTE_TO_LWORD(in);
END_FUNCTION

FUNCTION TO_LWORD__WORD : LWORD
    VAR_INPUT
        in : WORD;
    END_VAR

    TO_LWORD__WORD := WORD_TO_LWORD(in);
END_FUNCTION

FUNCTION TO_LWORD__DWORD : LWORD
    VAR_INPUT
        in : DWORD;
    END_VAR

    TO_LWORD__DWORD := DWORD_TO_LWORD(in);
END_FUNCTION

FUNCTION TO_LWORD__REAL : LWORD
    VAR_INPUT
        in : REAL;
    END_VAR

    TO_LWORD__REAL := REAL_TO_LWORD(in);
END_FUNCTION

FUNCTION TO_LWORD__LREAL : LWORD
    VAR_INPUT
        in : LREAL;
    END_VAR

    TO_LWORD__LREAL := LREAL_TO_LWORD(in);
END_FUNCTION

(* ---- to_date_time.st ---- *)
FUNCTION TO_TIME<T: ANY> : TIME
    VAR_INPUT
        in : T;
    END_VAR
END_FUNCTION

FUNCTION TO_TIME__TIME : TIME
    VAR_INPUT
        in : TIME;
    END_VAR

    TO_TIME__TIME := in;
END_FUNCTION

FUNCTION TO_TIME__LTIME : TIME
    VAR_INPUT
        in : LTIME;
    END_VAR

    TO_TIME__LTIME := LTIME_TO_TIME(in);
END_FUNCTION

FUNCTION TO_TIME__BOOL : TIME
    VAR_INPUT
        in : BOOL;
    END_VAR

    TO_TIME__BOOL := BOOL_TO_TIME(in);
END_FUNCTION

FUNCTION TO_TIME__BYTE : TIME
    VAR_INPUT
        in : BYTE;
    END_VAR

    TO_TIME__BYTE := BYTE_TO_TIME(in);
END_FUNCTION

FUNCTION TO_TIME__WORD : TIME
    VAR_INPUT
        in : WORD;
    END_VAR

    TO_TIME__WORD := WORD_TO_TIME(in);
END_FUNCTION

FUNCTION TO_TIME__DWORD : TIME
    VAR_INPUT
        in : DWORD;
    END_VAR

    TO_TIME__DWORD := DWORD_TO_TIME(in);
END_FUNCTION

FUNCTION TO_TIME__LWORD : TIME
    VAR_INPUT
        in : LWORD;
    END_VAR

    TO_TIME__LWORD := LWORD_TO_TIME(in);
END_FUNCTION

FUNCTION TO_TIME__SINT : TIME
    VAR_INPUT
        in : SINT;
    END_VAR

    TO_TIME__SINT := SINT_TO_TIME(in);
END_FUNCTION

FUNCTION TO_TIME__USINT : TIME
    VAR_INPUT
        in : USINT;
    END_VAR

    TO_TIME__USINT := USINT_TO_TIME(in);
END_FUNCTION

FUNCTION TO_TIME__INT : TIME
    VAR_INPUT
        in : INT;
    END_VAR

    TO_TIME__INT := INT_TO_TIME(in);
END_FUNCTION

FUNCTION TO_TIME__UINT : TIME
    VAR_INPUT
        in : UINT;
    END_VAR

    TO_TIME__UINT := UINT_TO_TIME(in);
END_FUNCTION

FUNCTION TO_TIME__DINT : TIME
    VAR_INPUT
        in : DINT;
    END_VAR

    TO_TIME__DINT := DINT_TO_TIME(in);
END_FUNCTION

FUNCTION TO_TIME__UDINT : TIME
    VAR_INPUT
        in : UDINT;
    END_VAR

    TO_TIME__UDINT := UDINT_TO_TIME(in);
END_FUNCTION

FUNCTION TO_TIME__LINT : TIME
    VAR_INPUT
        in : LINT;
    END_VAR

    TO_TIME__LINT := LINT_TO_TIME(in);
END_FUNCTION

FUNCTION TO_TIME__ULINT : TIME
    VAR_INPUT
        in : ULINT;
    END_VAR

    TO_TIME__ULINT := ULINT_TO_TIME(in);
END_FUNCTION

FUNCTION TO_TIME__REAL : TIME
    VAR_INPUT
        in : REAL;
    END_VAR

    TO_TIME__REAL := REAL_TO_TIME(in);
END_FUNCTION

FUNCTION TO_TIME__LREAL : TIME
    VAR_INPUT
        in : LREAL;
    END_VAR

    TO_TIME__LREAL := LREAL_TO_TIME(in);
END_FUNCTION

// -----------------------------------------------------------------------------------------------------------

FUNCTION TO_LTIME<T: ANY> : LTIME
    VAR_INPUT
        in : T;
    END_VAR
END_FUNCTION

FUNCTION TO_LTIME__LTIME : LTIME
    VAR_INPUT
        in : LTIME;
    END_VAR

    TO_LTIME__LTIME := in;
END_FUNCTION

FUNCTION TO_LTIME__TIME : LTIME
    VAR_INPUT
        in : TIME;
    END_VAR

    TO_LTIME__TIME := TIME_TO_LTIME(in);
END_FUNCTION

FUNCTION TO_LTIME__BOOL : LTIME
    VAR_INPUT
        in : BOOL;
    END_VAR

    TO_LTIME__BOOL := BOOL_TO_LTIME(in);
END_FUNCTION

FUNCTION TO_LTIME__BYTE : LTIME
    VAR_INPUT
        in : BYTE;
    END_VAR

    TO_LTIME__BYTE := BYTE_TO_LTIME(in);
END_FUNCTION

FUNCTION TO_LTIME__WORD : LTIME
    VAR_INPUT
        in : WORD;
    END_VAR

    TO_LTIME__WORD := WORD_TO_LTIME(in);
END_FUNCTION

FUNCTION TO_LTIME__DWORD : LTIME
    VAR_INPUT
        in : DWORD;
    END_VAR

    TO_LTIME__DWORD := DWORD_TO_LTIME(in);
END_FUNCTION

FUNCTION TO_LTIME__LWORD : LTIME
    VAR_INPUT
        in : LWORD;
    END_VAR

    TO_LTIME__LWORD := LWORD_TO_LTIME(in);
END_FUNCTION

FUNCTION TO_LTIME__SINT : LTIME
    VAR_INPUT
        in : SINT;
    END_VAR

    TO_LTIME__SINT := SINT_TO_LTIME(in);
END_FUNCTION

FUNCTION TO_LTIME__USINT : LTIME
    VAR_INPUT
        in : USINT;
    END_VAR

    TO_LTIME__USINT := USINT_TO_LTIME(in);
END_FUNCTION

FUNCTION TO_LTIME__INT : LTIME
    VAR_INPUT
        in : INT;
    END_VAR

    TO_LTIME__INT := INT_TO_LTIME(in);
END_FUNCTION

FUNCTION TO_LTIME__UINT : LTIME
    VAR_INPUT
        in : UINT;
    END_VAR

    TO_LTIME__UINT := UINT_TO_LTIME(in);
END_FUNCTION

FUNCTION TO_LTIME__DINT : LTIME
    VAR_INPUT
        in : DINT;
    END_VAR

    TO_LTIME__DINT := DINT_TO_LTIME(in);
END_FUNCTION

FUNCTION TO_LTIME__UDINT : LTIME
    VAR_INPUT
        in : UDINT;
    END_VAR

    TO_LTIME__UDINT := UDINT_TO_LTIME(in);
END_FUNCTION

FUNCTION TO_LTIME__LINT : LTIME
    VAR_INPUT
        in : LINT;
    END_VAR

    TO_LTIME__LINT := LINT_TO_LTIME(in);
END_FUNCTION

FUNCTION TO_LTIME__ULINT : LTIME
    VAR_INPUT
        in : ULINT;
    END_VAR

    TO_LTIME__ULINT := ULINT_TO_LTIME(in);
END_FUNCTION

FUNCTION TO_LTIME__REAL : LTIME
    VAR_INPUT
        in : REAL;
    END_VAR

    TO_LTIME__REAL := REAL_TO_LTIME(in);
END_FUNCTION

FUNCTION TO_LTIME__LREAL : LTIME
    VAR_INPUT
        in : LREAL;
    END_VAR

    TO_LTIME__LREAL := LREAL_TO_LTIME(in);
END_FUNCTION

// -----------------------------------------------------------------------------------------------------------

FUNCTION TO_DT<T: ANY> : DT
    VAR_INPUT
        in : T;
    END_VAR
END_FUNCTION

FUNCTION TO_DT__DATE_AND_TIME : DT
    VAR_INPUT
        in : DT;
    END_VAR

    TO_DT__DATE_AND_TIME := in;
END_FUNCTION

FUNCTION TO_DT__LDATE_AND_TIME : DT
    VAR_INPUT
        in : LDT;
    END_VAR

    TO_DT__LDATE_AND_TIME := LDT_TO_DT(in);
END_FUNCTION

// -----------------------------------------------------------------------------------------------------------

FUNCTION TO_DATE<T: ANY> : DATE
    VAR_INPUT
        in : T;
    END_VAR
END_FUNCTION

FUNCTION TO_DATE__DATE_AND_TIME : DATE
    VAR_INPUT
        in : DT;
    END_VAR

    TO_DATE__DATE_AND_TIME := DT_TO_DATE(in);
END_FUNCTION

FUNCTION TO_DATE__LDATE_AND_TIME : DATE
    VAR_INPUT
        in : LDT;
    END_VAR

    TO_DATE__LDATE_AND_TIME := LDT_TO_DATE(in);
END_FUNCTION

// -----------------------------------------------------------------------------------------------------------

FUNCTION TO_LDATE<T: ANY> : LDATE
    VAR_INPUT
        in : T;
    END_VAR
END_FUNCTION

FUNCTION TO_LDATE__DATE_AND_TIME : LDATE
    VAR_INPUT
        in : DT;
    END_VAR

    TO_LDATE__DATE_AND_TIME := DT_TO_LDATE(in);
END_FUNCTION

FUNCTION TO_LDATE__LDATE_AND_TIME : LDATE
    VAR_INPUT
        in : LDT;
    END_VAR

    TO_LDATE__LDATE_AND_TIME := LDATE_AND_TIME_TO_LDATE(in);
END_FUNCTION

// -----------------------------------------------------------------------------------------------------------

FUNCTION TO_TOD<T: ANY> : TOD
    VAR_INPUT
        in : T;
    END_VAR
END_FUNCTION

FUNCTION TO_TOD__DATE_AND_TIME : TOD
    VAR_INPUT
        in : DT;
    END_VAR

    TO_TOD__DATE_AND_TIME := DT_TO_TOD(in);
END_FUNCTION

FUNCTION TO_TOD__LDATE_AND_TIME : TOD
    VAR_INPUT
        in : LDT;
    END_VAR

    TO_TOD__LDATE_AND_TIME := LDT_TO_TOD(in);
END_FUNCTION

FUNCTION TO_TOD__TIME_OF_DAY : TOD
    VAR_INPUT
        in : TOD;
    END_VAR

    TO_TOD__TIME_OF_DAY := in;
END_FUNCTION

FUNCTION TO_TOD__LTIME_OF_DAY : TOD
    VAR_INPUT
        in : LTOD;
    END_VAR

    TO_TOD__LTIME_OF_DAY := LTOD_TO_TOD(in);
END_FUNCTION

// -----------------------------------------------------------------------------------------------------------

FUNCTION TO_LTOD<T: ANY> : LTOD
    VAR_INPUT
        in : T;
    END_VAR
END_FUNCTION

FUNCTION TO_LTOD__DATE_AND_TIME : LTOD
    VAR_INPUT
        in : DT;
    END_VAR

    TO_LTOD__DATE_AND_TIME := DT_TO_LTOD(in);
END_FUNCTION

FUNCTION TO_LTOD__LDATE_AND_TIME : LTOD
    VAR_INPUT
        in : LDT;
    END_VAR

    TO_LTOD__LDATE_AND_TIME := LDT_TO_LTOD(in);
END_FUNCTION

FUNCTION TO_LTOD__TIME_OF_DAY : LTOD
    VAR_INPUT
        in : TOD;
    END_VAR

    TO_LTOD__TIME_OF_DAY := TOD_TO_LTOD(in);
END_FUNCTION

FUNCTION TO_LTOD__LTIME_OF_DAY : LTOD
    VAR_INPUT
        in : LTOD;
    END_VAR

    TO_LTOD__LTIME_OF_DAY := in;
END_FUNCTION

// -----------------------------------------------------------------------------------------------------------

FUNCTION TO_LDT<T: ANY> : LDT
    VAR_INPUT
        in : T;
    END_VAR
END_FUNCTION

FUNCTION TO_LDT__DATE_AND_TIME : LDT
    VAR_INPUT
        in : DT;
    END_VAR

    TO_LDT__DATE_AND_TIME := DT_TO_LDT(in);
END_FUNCTION

FUNCTION TO_LDT__LDATE_AND_TIME : LDT
    VAR_INPUT
        in : LDT;
    END_VAR

    TO_LDT__LDATE_AND_TIME := in;
END_FUNCTION

(* ---- to_num.st ---- *)
(********************
*
* Converts any other numerical value to SINT
*
*********************)
FUNCTION TO_SINT<T: ANY_NUM> : SINT
    VAR_INPUT
        in : T;
    END_VAR
END_FUNCTION

(********************
*
* Converts SINT to SINT
*
*********************)
FUNCTION TO_SINT__SINT : SINT
    VAR_INPUT
        in : SINT;
    END_VAR

    TO_SINT__SINT := in;
END_FUNCTION

(********************
*
* Converts SINT to USINT
*
*********************)
FUNCTION TO_USINT__SINT : USINT
    VAR_INPUT
        in : SINT;
    END_VAR

    TO_USINT__SINT := SINT_TO_USINT(in);
END_FUNCTION

(********************
*
* Converts SINT to INT
*
*********************)
FUNCTION TO_INT__SINT : INT
    VAR_INPUT
        in : SINT;
    END_VAR

    TO_INT__SINT := SINT_TO_INT(in);
END_FUNCTION

(********************
*
* Converts SINT to UINT
*
*********************)
FUNCTION TO_UINT__SINT : UINT
    VAR_INPUT
        in : SINT;
    END_VAR

    TO_UINT__SINT := SINT_TO_UINT(in);
END_FUNCTION

(********************
*
* Converts SINT to DINT
*
*********************)
FUNCTION TO_DINT__SINT : DINT
    VAR_INPUT
        in : SINT;
    END_VAR

    TO_DINT__SINT := SINT_TO_DINT(in);
END_FUNCTION

(********************
*
* Converts SINT to UDINT
*
*********************)
FUNCTION TO_UDINT__SINT : UDINT
    VAR_INPUT
        in : SINT;
    END_VAR

    TO_UDINT__SINT := SINT_TO_UDINT(in);
END_FUNCTION

(********************
*
* Converts SINT to LINT
*
*********************)
FUNCTION TO_LINT__SINT : LINT
    VAR_INPUT
        in : SINT;
    END_VAR

    TO_LINT__SINT := SINT_TO_LINT(in);
END_FUNCTION

(********************
*
* Converts SINT to ULINT
*
*********************)
FUNCTION TO_ULINT__SINT : ULINT
    VAR_INPUT
        in : SINT;
    END_VAR

    TO_ULINT__SINT := SINT_TO_ULINT(in);
END_FUNCTION

(********************
*
* Converts SINT to REAL
*
*********************)
FUNCTION TO_REAL__SINT : REAL
    VAR_INPUT
        in : SINT;
    END_VAR

    TO_REAL__SINT := SINT_TO_REAL(in);
END_FUNCTION

(********************
*
* Converts SINT to LREAL
*
*********************)
FUNCTION TO_LREAL__SINT : LREAL
    VAR_INPUT
        in : SINT;
    END_VAR

    TO_LREAL__SINT := SINT_TO_LREAL(in);
END_FUNCTION

(********************
*
* Converts any other numerical value to USINT
*
*********************)
FUNCTION TO_USINT<T: ANY_NUM> : USINT
    VAR_INPUT
        in : T;
    END_VAR
END_FUNCTION

(********************
*
* Converts USINT to SINT
*
*********************)
FUNCTION TO_SINT__USINT : SINT
    VAR_INPUT
        in : USINT;
    END_VAR

    TO_SINT__USINT := USINT_TO_SINT(in);
END_FUNCTION

(********************
*
* Converts USINT to USINT
*
*********************)
FUNCTION TO_USINT__USINT : USINT
    VAR_INPUT
        in : USINT;
    END_VAR

    TO_USINT__USINT := in;
END_FUNCTION

(********************
*
* Converts USINT to INT
*
*********************)
FUNCTION TO_INT__USINT : INT
    VAR_INPUT
        in : USINT;
    END_VAR

    TO_INT__USINT := USINT_TO_INT(in);
END_FUNCTION

(********************
*
* Converts USINT to UINT
*
*********************)
FUNCTION TO_UINT__USINT : UINT
    VAR_INPUT
        in : USINT;
    END_VAR

    TO_UINT__USINT := USINT_TO_UINT(in);
END_FUNCTION

(********************
*
* Converts USINT to DINT
*
*********************)
FUNCTION TO_DINT__USINT : DINT
    VAR_INPUT
        in : USINT;
    END_VAR

    TO_DINT__USINT := USINT_TO_DINT(in);
END_FUNCTION

(********************
*
* Converts USINT to UDINT
*
*********************)
FUNCTION TO_UDINT__USINT : UDINT
    VAR_INPUT
        in : USINT;
    END_VAR

    TO_UDINT__USINT := USINT_TO_UDINT(in);
END_FUNCTION

(********************
*
* Converts USINT to LINT
*
*********************)
FUNCTION TO_LINT__USINT : LINT
    VAR_INPUT
        in : USINT;
    END_VAR

    TO_LINT__USINT := USINT_TO_LINT(in);
END_FUNCTION

(********************
*
* Converts USINT to ULINT
*
*********************)
FUNCTION TO_ULINT__USINT : ULINT
    VAR_INPUT
        in : USINT;
    END_VAR

    TO_ULINT__USINT := USINT_TO_ULINT(in);
END_FUNCTION

(********************
*
* Converts USINT to REAL
*
*********************)
FUNCTION TO_REAL__USINT : REAL
    VAR_INPUT
        in : USINT;
    END_VAR

    TO_REAL__USINT := USINT_TO_REAL(in);
END_FUNCTION

(********************
*
* Converts USINT to LREAL
*
*********************)
FUNCTION TO_LREAL__USINT : LREAL
    VAR_INPUT
        in : USINT;
    END_VAR

    TO_LREAL__USINT := USINT_TO_LREAL(in);
END_FUNCTION

(********************
*
* Converts any other numerical value to INT
*
*********************)
FUNCTION TO_INT<T: ANY_NUM> : INT
    VAR_INPUT
        in : T;
    END_VAR
END_FUNCTION

(********************
*
* Converts INT to SINT
*
*********************)
FUNCTION TO_SINT__INT : SINT
    VAR_INPUT
        in : INT;
    END_VAR

    TO_SINT__INT := INT_TO_SINT(in);
END_FUNCTION

(********************
*
* Converts INT to USINT
*
*********************)
FUNCTION TO_USINT__INT : USINT
    VAR_INPUT
        in : INT;
    END_VAR

    TO_USINT__INT := INT_TO_USINT(in);
END_FUNCTION

(********************
*
* Converts INT to INT
*
*********************)
FUNCTION TO_INT__INT : INT
    VAR_INPUT
        in : INT;
    END_VAR

    TO_INT__INT := in;
END_FUNCTION

(********************
*
* Converts INT to UINT
*
*********************)
FUNCTION TO_UINT__INT : UINT
    VAR_INPUT
        in : INT;
    END_VAR

    TO_UINT__INT := INT_TO_UINT(in);
END_FUNCTION

(********************
*
* Converts INT to DINT
*
*********************)
FUNCTION TO_DINT__INT : DINT
    VAR_INPUT
        in : INT;
    END_VAR

    TO_DINT__INT := INT_TO_DINT(in);
END_FUNCTION

(********************
*
* Converts INT to UDINT
*
*********************)
FUNCTION TO_UDINT__INT : UDINT
    VAR_INPUT
        in : INT;
    END_VAR

    TO_UDINT__INT := INT_TO_UDINT(in);
END_FUNCTION

(********************
*
* Converts INT to LINT
*
*********************)
FUNCTION TO_LINT__INT : LINT
    VAR_INPUT
        in : INT;
    END_VAR

    TO_LINT__INT := INT_TO_LINT(in);
END_FUNCTION

(********************
*
* Converts INT to ULINT
*
*********************)
FUNCTION TO_ULINT__INT : ULINT
    VAR_INPUT
        in : INT;
    END_VAR

    TO_ULINT__INT := INT_TO_ULINT(in);
END_FUNCTION

(********************
*
* Converts INT to REAL
*
*********************)
FUNCTION TO_REAL__INT : REAL
    VAR_INPUT
        in : INT;
    END_VAR

    TO_REAL__INT := INT_TO_REAL(in);
END_FUNCTION

(********************
*
* Converts INT to LREAL
*
*********************)
FUNCTION TO_LREAL__INT : LREAL
    VAR_INPUT
        in : INT;
    END_VAR

    TO_LREAL__INT := INT_TO_LREAL(in);
END_FUNCTION

(********************
*
* Converts any other numerical value to UINT
*
*********************)
FUNCTION TO_UINT<T: ANY_NUM> : UINT
    VAR_INPUT
        in : T;
    END_VAR
END_FUNCTION

(********************
*
* Converts UINT to SINT
*
*********************)
FUNCTION TO_SINT__UINT : SINT
    VAR_INPUT
        in : UINT;
    END_VAR

    TO_SINT__UINT := UINT_TO_SINT(in);
END_FUNCTION

(********************
*
* Converts UINT to USINT
*
*********************)
FUNCTION TO_USINT__UINT : USINT
    VAR_INPUT
        in : UINT;
    END_VAR

    TO_USINT__UINT := UINT_TO_USINT(in);
END_FUNCTION

(********************
*
* Converts UINT to INT
*
*********************)
FUNCTION TO_INT__UINT : INT
    VAR_INPUT
        in : UINT;
    END_VAR

    TO_INT__UINT := UINT_TO_INT(in);
END_FUNCTION

(********************
*
* Converts UINT to UINT
*
*********************)
FUNCTION TO_UINT__UINT : UINT
    VAR_INPUT
        in : UINT;
    END_VAR

    TO_UINT__UINT := in;
END_FUNCTION

(********************
*
* Converts UINT to DINT
*
*********************)
FUNCTION TO_DINT__UINT : DINT
    VAR_INPUT
        in : UINT;
    END_VAR

    TO_DINT__UINT := UINT_TO_DINT(in);
END_FUNCTION

(********************
*
* Converts UINT to UDINT
*
*********************)
FUNCTION TO_UDINT__UINT : UDINT
    VAR_INPUT
        in : UINT;
    END_VAR

    TO_UDINT__UINT := UINT_TO_UDINT(in);
END_FUNCTION

(********************
*
* Converts UINT to LINT
*
*********************)
FUNCTION TO_LINT__UINT : LINT
    VAR_INPUT
        in : UINT;
    END_VAR

    TO_LINT__UINT := UINT_TO_LINT(in);
END_FUNCTION

(********************
*
* Converts UINT to ULINT
*
*********************)
FUNCTION TO_ULINT__UINT : ULINT
    VAR_INPUT
        in : UINT;
    END_VAR

    TO_ULINT__UINT := UINT_TO_ULINT(in);
END_FUNCTION

(********************
*
* Converts UINT to REAL
*
*********************)
FUNCTION TO_REAL__UINT : REAL
    VAR_INPUT
        in : UINT;
    END_VAR

    TO_REAL__UINT := UINT_TO_REAL(in);
END_FUNCTION

(********************
*
* Converts UINT to LREAL
*
*********************)
FUNCTION TO_LREAL__UINT : LREAL
    VAR_INPUT
        in : UINT;
    END_VAR

    TO_LREAL__UINT := UINT_TO_LREAL(in);
END_FUNCTION

(********************
*
* Converts any other numerical value to DINT
*
*********************)
FUNCTION TO_DINT<T: ANY_NUM> : DINT
    VAR_INPUT
        in : T;
    END_VAR
END_FUNCTION

(********************
*
* Converts DINT to SINT
*
*********************)
FUNCTION TO_SINT__DINT : SINT
    VAR_INPUT
        in : DINT;
    END_VAR

    TO_SINT__DINT := DINT_TO_SINT(in);
END_FUNCTION

(********************
*
* Converts DINT to USINT
*
*********************)
FUNCTION TO_USINT__DINT : USINT
    VAR_INPUT
        in : DINT;
    END_VAR

    TO_USINT__DINT := DINT_TO_USINT(in);
END_FUNCTION

(********************
*
* Converts DINT to INT
*
*********************)
FUNCTION TO_INT__DINT : INT
    VAR_INPUT
        in : DINT;
    END_VAR

    TO_INT__DINT := DINT_TO_INT(in);
END_FUNCTION

(********************
*
* Converts DINT to UINT
*
*********************)
FUNCTION TO_UINT__DINT : UINT
    VAR_INPUT
        in : DINT;
    END_VAR

    TO_UINT__DINT := DINT_TO_UINT(in);
END_FUNCTION

(********************
*
* Converts DINT to DINT
*
*********************)
FUNCTION TO_DINT__DINT : DINT
    VAR_INPUT
        in : DINT;
    END_VAR

    TO_DINT__DINT := in;
END_FUNCTION

(********************
*
* Converts DINT to UDINT
*
*********************)
FUNCTION TO_UDINT__DINT : UDINT
    VAR_INPUT
        in : DINT;
    END_VAR

    TO_UDINT__DINT := DINT_TO_UDINT(in);
END_FUNCTION

(********************
*
* Converts DINT to LINT
*
*********************)
FUNCTION TO_LINT__DINT : LINT
    VAR_INPUT
        in : DINT;
    END_VAR

    TO_LINT__DINT := DINT_TO_LINT(in);
END_FUNCTION

(********************
*
* Converts DINT to ULINT
*
*********************)
FUNCTION TO_ULINT__DINT : ULINT
    VAR_INPUT
        in : DINT;
    END_VAR

    TO_ULINT__DINT := DINT_TO_ULINT(in);
END_FUNCTION

(********************
*
* Converts DINT to REAL
*
*********************)
FUNCTION TO_REAL__DINT : REAL
    VAR_INPUT
        in : DINT;
    END_VAR

    TO_REAL__DINT := DINT_TO_REAL(in);
END_FUNCTION

(********************
*
* Converts DINT to LREAL
*
*********************)
FUNCTION TO_LREAL__DINT : LREAL
    VAR_INPUT
        in : DINT;
    END_VAR

    TO_LREAL__DINT := DINT_TO_LREAL(in);
END_FUNCTION

(********************
*
* Converts any other numerical value to UDINT
*
*********************)
FUNCTION TO_UDINT<T: ANY_NUM> : UDINT
    VAR_INPUT
        in : T;
    END_VAR
END_FUNCTION

(********************
*
* Converts UDINT to SINT
*
*********************)
FUNCTION TO_SINT__UDINT : SINT
    VAR_INPUT
        in : UDINT;
    END_VAR

    TO_SINT__UDINT := UDINT_TO_SINT(in);
END_FUNCTION

(********************
*
* Converts UDINT to USINT
*
*********************)
FUNCTION TO_USINT__UDINT : USINT
    VAR_INPUT
        in : UDINT;
    END_VAR

    TO_USINT__UDINT := UDINT_TO_USINT(in);
END_FUNCTION

(********************
*
* Converts UDINT to INT
*
*********************)
FUNCTION TO_INT__UDINT : INT
    VAR_INPUT
        in : UDINT;
    END_VAR

    TO_INT__UDINT := UDINT_TO_INT(in);
END_FUNCTION

(********************
*
* Converts UDINT to UINT
*
*********************)
FUNCTION TO_UINT__UDINT : UINT
    VAR_INPUT
        in : UDINT;
    END_VAR

    TO_UINT__UDINT := UDINT_TO_UINT(in);
END_FUNCTION

(********************
*
* Converts UDINT to DINT
*
*********************)
FUNCTION TO_DINT__UDINT : DINT
    VAR_INPUT
        in : UDINT;
    END_VAR

    TO_DINT__UDINT := UDINT_TO_DINT(in);
END_FUNCTION

(********************
*
* Converts UDINT to UDINT
*
*********************)
FUNCTION TO_UDINT__UDINT : UDINT
    VAR_INPUT
        in : UDINT;
    END_VAR

    TO_UDINT__UDINT := in;
END_FUNCTION

(********************
*
* Converts UDINT to LINT
*
*********************)
FUNCTION TO_LINT__UDINT : LINT
    VAR_INPUT
        in : UDINT;
    END_VAR

    TO_LINT__UDINT := UDINT_TO_LINT(in);
END_FUNCTION

(********************
*
* Converts UDINT to ULINT
*
*********************)
FUNCTION TO_ULINT__UDINT : ULINT
    VAR_INPUT
        in : UDINT;
    END_VAR

    TO_ULINT__UDINT := UDINT_TO_ULINT(in);
END_FUNCTION

(********************
*
* Converts UDINT to REAL
*
*********************)
FUNCTION TO_REAL__UDINT : REAL
    VAR_INPUT
        in : UDINT;
    END_VAR

    TO_REAL__UDINT := UDINT_TO_REAL(in);
END_FUNCTION

(********************
*
* Converts UDINT to LREAL
*
*********************)
FUNCTION TO_LREAL__UDINT : LREAL
    VAR_INPUT
        in : UDINT;
    END_VAR

    TO_LREAL__UDINT := UDINT_TO_LREAL(in);
END_FUNCTION

(********************
*
* Converts any other numerical value to LINT
*
*********************)
FUNCTION TO_LINT<T: ANY_NUM> : LINT
    VAR_INPUT
        in : T;
    END_VAR
END_FUNCTION

(********************
*
* Converts LINT to SINT
*
*********************)
FUNCTION TO_SINT__LINT : SINT
    VAR_INPUT
        in : LINT;
    END_VAR

    TO_SINT__LINT := LINT_TO_SINT(in);
END_FUNCTION

(********************
*
* Converts LINT to USINT
*
*********************)
FUNCTION TO_USINT__LINT : USINT
    VAR_INPUT
        in : LINT;
    END_VAR

    TO_USINT__LINT := LINT_TO_USINT(in);
END_FUNCTION

(********************
*
* Converts LINT to INT
*
*********************)
FUNCTION TO_INT__LINT : INT
    VAR_INPUT
        in : LINT;
    END_VAR

    TO_INT__LINT := LINT_TO_INT(in);
END_FUNCTION

(********************
*
* Converts LINT to UINT
*
*********************)
FUNCTION TO_UINT__LINT : UINT
    VAR_INPUT
        in : LINT;
    END_VAR

    TO_UINT__LINT := LINT_TO_UINT(in);
END_FUNCTION

(********************
*
* Converts LINT to DINT
*
*********************)
FUNCTION TO_DINT__LINT : DINT
    VAR_INPUT
        in : LINT;
    END_VAR

    TO_DINT__LINT := LINT_TO_DINT(in);
END_FUNCTION

(********************
*
* Converts LINT to UDINT
*
*********************)
FUNCTION TO_UDINT__LINT : UDINT
    VAR_INPUT
        in : LINT;
    END_VAR

    TO_UDINT__LINT := LINT_TO_UDINT(in);
END_FUNCTION

(********************
*
* Converts LINT to LINT
*
*********************)
FUNCTION TO_LINT__LINT : LINT
    VAR_INPUT
        in : LINT;
    END_VAR

    TO_LINT__LINT := in;
END_FUNCTION

(********************
*
* Converts LINT to ULINT
*
*********************)
FUNCTION TO_ULINT__LINT : ULINT
    VAR_INPUT
        in : LINT;
    END_VAR

    TO_ULINT__LINT := LINT_TO_ULINT(in);
END_FUNCTION

(********************
*
* Converts LINT to REAL
*
*********************)
FUNCTION TO_REAL__LINT : REAL
    VAR_INPUT
        in : LINT;
    END_VAR

    TO_REAL__LINT := LINT_TO_REAL(in);
END_FUNCTION

(********************
*
* Converts LINT to LREAL
*
*********************)
FUNCTION TO_LREAL__LINT : LREAL
    VAR_INPUT
        in : LINT;
    END_VAR

    TO_LREAL__LINT := LINT_TO_LREAL(in);
END_FUNCTION

(********************
*
* Converts any other numerical value to ULINT
*
*********************)
FUNCTION TO_ULINT<T: ANY_NUM> : ULINT
    VAR_INPUT
        in : T;
    END_VAR
END_FUNCTION

(********************
*
* Converts ULINT to SINT
*
*********************)
FUNCTION TO_SINT__ULINT : SINT
    VAR_INPUT
        in : ULINT;
    END_VAR

    TO_SINT__ULINT := ULINT_TO_SINT(in);
END_FUNCTION

(********************
*
* Converts ULINT to USINT
*
*********************)
FUNCTION TO_USINT__ULINT : USINT
    VAR_INPUT
        in : ULINT;
    END_VAR

    TO_USINT__ULINT := ULINT_TO_USINT(in);
END_FUNCTION

(********************
*
* Converts ULINT to INT
*
*********************)
FUNCTION TO_INT__ULINT : INT
    VAR_INPUT
        in : ULINT;
    END_VAR

    TO_INT__ULINT := ULINT_TO_INT(in);
END_FUNCTION

(********************
*
* Converts ULINT to UINT
*
*********************)
FUNCTION TO_UINT__ULINT : UINT
    VAR_INPUT
        in : ULINT;
    END_VAR

    TO_UINT__ULINT := ULINT_TO_UINT(in);
END_FUNCTION

(********************
*
* Converts ULINT to DINT
*
*********************)
FUNCTION TO_DINT__ULINT : DINT
    VAR_INPUT
        in : ULINT;
    END_VAR

    TO_DINT__ULINT := ULINT_TO_DINT(in);
END_FUNCTION

(********************
*
* Converts ULINT to UDINT
*
*********************)
FUNCTION TO_UDINT__ULINT : UDINT
    VAR_INPUT
        in : ULINT;
    END_VAR

    TO_UDINT__ULINT := ULINT_TO_UDINT(in);
END_FUNCTION

(********************
*
* Converts ULINT to LINT
*
*********************)
FUNCTION TO_LINT__ULINT : LINT
    VAR_INPUT
        in : ULINT;
    END_VAR

    TO_LINT__ULINT := ULINT_TO_LINT(in);
END_FUNCTION

(********************
*
* Converts ULINT to ULINT
*
*********************)
FUNCTION TO_ULINT__ULINT : ULINT
    VAR_INPUT
        in : ULINT;
    END_VAR

    TO_ULINT__ULINT := in;
END_FUNCTION

(********************
*
* Converts ULINT to REAL
*
*********************)
FUNCTION TO_REAL__ULINT : REAL
    VAR_INPUT
        in : ULINT;
    END_VAR

    TO_REAL__ULINT := ULINT_TO_REAL(in);
END_FUNCTION

(********************
*
* Converts ULINT to LREAL
*
*********************)
FUNCTION TO_LREAL__ULINT : LREAL
    VAR_INPUT
        in : ULINT;
    END_VAR

    TO_LREAL__ULINT := ULINT_TO_LREAL(in);
END_FUNCTION

(********************
*
* Converts any other numerical value to REAL
*
*********************)
FUNCTION TO_REAL<T: ANY_NUM> : REAL
    VAR_INPUT
        in : T;
    END_VAR
END_FUNCTION

(********************
*
* Converts REAL to SINT
*
*********************)
FUNCTION TO_SINT__REAL : SINT
    VAR_INPUT
        in : REAL;
    END_VAR

    TO_SINT__REAL := REAL_TO_SINT(in);
END_FUNCTION

(********************
*
* Converts REAL to USINT
*
*********************)
FUNCTION TO_USINT__REAL : USINT
    VAR_INPUT
        in : REAL;
    END_VAR

    TO_USINT__REAL := REAL_TO_USINT(in);
END_FUNCTION

(********************
*
* Converts REAL to INT
*
*********************)
FUNCTION TO_INT__REAL : INT
    VAR_INPUT
        in : REAL;
    END_VAR

    TO_INT__REAL := REAL_TO_INT(in);
END_FUNCTION

(********************
*
* Converts REAL to UINT
*
*********************)
FUNCTION TO_UINT__REAL : UINT
    VAR_INPUT
        in : REAL;
    END_VAR

    TO_UINT__REAL := REAL_TO_UINT(in);
END_FUNCTION

(********************
*
* Converts REAL to DINT
*
*********************)
FUNCTION TO_DINT__REAL : DINT
    VAR_INPUT
        in : REAL;
    END_VAR

    TO_DINT__REAL := REAL_TO_DINT(in);
END_FUNCTION

(********************
*
* Converts REAL to UDINT
*
*********************)
FUNCTION TO_UDINT__REAL : UDINT
    VAR_INPUT
        in : REAL;
    END_VAR

    TO_UDINT__REAL := REAL_TO_UDINT(in);
END_FUNCTION

(********************
*
* Converts REAL to LINT
*
*********************)
FUNCTION TO_LINT__REAL : LINT
    VAR_INPUT
        in : REAL;
    END_VAR

    TO_LINT__REAL := REAL_TO_LINT(in);
END_FUNCTION

(********************
*
* Converts REAL to ULINT
*
*********************)
FUNCTION TO_ULINT__REAL : ULINT
    VAR_INPUT
        in : REAL;
    END_VAR

    TO_ULINT__REAL := REAL_TO_ULINT(in);
END_FUNCTION

(********************
*
* Converts REAL to REAL
*
*********************)
FUNCTION TO_REAL__REAL : REAL
    VAR_INPUT
        in : REAL;
    END_VAR

    TO_REAL__REAL := in;
END_FUNCTION

(********************
*
* Converts REAL to LREAL
*
*********************)
FUNCTION TO_LREAL__REAL : LREAL
    VAR_INPUT
        in : REAL;
    END_VAR

    TO_LREAL__REAL := REAL_TO_LREAL(in);
END_FUNCTION

(********************
*
* Converts any other numerical value to LREAL
*
*********************)
FUNCTION TO_LREAL<T: ANY_NUM> : LREAL
    VAR_INPUT
        in : T;
    END_VAR
END_FUNCTION

(********************
*
* Converts LREAL to SINT
*
*********************)
FUNCTION TO_SINT__LREAL : SINT
    VAR_INPUT
        in : LREAL;
    END_VAR

    TO_SINT__LREAL := LREAL_TO_SINT(in);
END_FUNCTION

(********************
*
* Converts LREAL to USINT
*
*********************)
FUNCTION TO_USINT__LREAL : USINT
    VAR_INPUT
        in : LREAL;
    END_VAR

    TO_USINT__LREAL := LREAL_TO_USINT(in);
END_FUNCTION

(********************
*
* Converts LREAL to INT
*
*********************)
FUNCTION TO_INT__LREAL : INT
    VAR_INPUT
        in : LREAL;
    END_VAR

    TO_INT__LREAL := LREAL_TO_INT(in);
END_FUNCTION

(********************
*
* Converts LREAL to UINT
*
*********************)
FUNCTION TO_UINT__LREAL : UINT
    VAR_INPUT
        in : LREAL;
    END_VAR

    TO_UINT__LREAL := LREAL_TO_UINT(in);
END_FUNCTION

(********************
*
* Converts LREAL to DINT
*
*********************)
FUNCTION TO_DINT__LREAL : DINT
    VAR_INPUT
        in : LREAL;
    END_VAR

    TO_DINT__LREAL := LREAL_TO_DINT(in);
END_FUNCTION

(********************
*
* Converts LREAL to UDINT
*
*********************)
FUNCTION TO_UDINT__LREAL : UDINT
    VAR_INPUT
        in : LREAL;
    END_VAR

    TO_UDINT__LREAL := LREAL_TO_UDINT(in);
END_FUNCTION

(********************
*
* Converts LREAL to LINT
*
*********************)
FUNCTION TO_LINT__LREAL : LINT
    VAR_INPUT
        in : LREAL;
    END_VAR

    TO_LINT__LREAL := LREAL_TO_LINT(in);
END_FUNCTION

(********************
*
* Converts LREAL to ULINT
*
*********************)
FUNCTION TO_ULINT__LREAL : ULINT
    VAR_INPUT
        in : LREAL;
    END_VAR

    TO_ULINT__LREAL := LREAL_TO_ULINT(in);
END_FUNCTION

(********************
*
* Converts LREAL to REAL
*
*********************)
FUNCTION TO_REAL__LREAL : REAL
    VAR_INPUT
        in : LREAL;
    END_VAR

    TO_REAL__LREAL := LREAL_TO_REAL(in);
END_FUNCTION

(********************
*
* Converts LREAL to LREAL
*
*********************)
FUNCTION TO_LREAL__LREAL : LREAL
    VAR_INPUT
        in : LREAL;
    END_VAR

    TO_LREAL__LREAL := in;
END_FUNCTION

(* ---- to_string.st ---- *)
FUNCTION TO_CHAR<T: ANY> : CHAR
    VAR_INPUT
        in : T;
    END_VAR
END_FUNCTION

FUNCTION TO_CHAR__CHAR : CHAR
    VAR_INPUT
        in : CHAR;
    END_VAR

    TO_CHAR__CHAR := in;
END_FUNCTION

FUNCTION TO_CHAR__WCHAR : CHAR
    VAR_INPUT
        in : WCHAR;
    END_VAR

    TO_CHAR__WCHAR := WCHAR_TO_CHAR(in);
END_FUNCTION

FUNCTION TO_CHAR__STRING : CHAR
    VAR_INPUT {ref}
        in : STRING;
    END_VAR

    TO_CHAR__STRING := STRING_TO_CHAR(in);
END_FUNCTION

// -----------------------------------------------------------------------------------------------------------

FUNCTION TO_WCHAR<T: ANY> : WCHAR
    VAR_INPUT
        in : T;
    END_VAR
END_FUNCTION

FUNCTION TO_WCHAR__WCHAR : WCHAR
    VAR_INPUT
        in : WCHAR;
    END_VAR

    TO_WCHAR__WCHAR := in;
END_FUNCTION

FUNCTION TO_WCHAR__CHAR : WCHAR
    VAR_INPUT
        in : CHAR;
    END_VAR

    TO_WCHAR__CHAR := CHAR_TO_WCHAR(in);

END_FUNCTION

FUNCTION TO_WCHAR__WSTRING : WCHAR
    VAR_INPUT {ref}
        in : WSTRING;
    END_VAR

    TO_WCHAR__WSTRING := WSTRING_TO_WCHAR(in);
END_FUNCTION

// -----------------------------------------------------------------------------------------------------------

FUNCTION TO_STRING<T: ANY> : STRING[__STRING_LENGTH]
    VAR_INPUT
        in : T;
    END_VAR
END_FUNCTION

FUNCTION TO_STRING__STRING : STRING[__STRING_LENGTH]
    VAR_INPUT {ref}
        in : STRING;
    END_VAR

    TO_STRING__STRING := in;
END_FUNCTION

FUNCTION TO_STRING__CHAR : STRING
    VAR_INPUT
        in : CHAR;
    END_VAR

    TO_STRING__CHAR := CHAR_TO_STRING(in);
END_FUNCTION

FUNCTION TO_STRING__WSTRING : STRING[__STRING_LENGTH]
    VAR_INPUT {ref}
        in : WSTRING;
    END_VAR

    WSTRING_TO_STRING_EXT(in, TO_STRING__WSTRING);
END_FUNCTION

// Numeric, bit-string and date/time monomorphizations of the generic TO_STRING, each
// delegating to the corresponding typed <T>_TO_STRING conversion function.

FUNCTION TO_STRING__DINT : STRING[__STRING_LENGTH]
    VAR_INPUT
        in : DINT;
    END_VAR

    TO_STRING__DINT := DINT_TO_STRING(in);
END_FUNCTION

FUNCTION TO_STRING__LINT : STRING[__STRING_LENGTH]
    VAR_INPUT
        in : LINT;
    END_VAR

    TO_STRING__LINT := LINT_TO_STRING(in);
END_FUNCTION

FUNCTION TO_STRING__USINT : STRING[__STRING_LENGTH]
    VAR_INPUT
        in : USINT;
    END_VAR

    TO_STRING__USINT := USINT_TO_STRING(in);
END_FUNCTION

FUNCTION TO_STRING__UINT : STRING[__STRING_LENGTH]
    VAR_INPUT
        in : UINT;
    END_VAR

    TO_STRING__UINT := UINT_TO_STRING(in);
END_FUNCTION

FUNCTION TO_STRING__UDINT : STRING[__STRING_LENGTH]
    VAR_INPUT
        in : UDINT;
    END_VAR

    TO_STRING__UDINT := UDINT_TO_STRING(in);
END_FUNCTION

FUNCTION TO_STRING__ULINT : STRING[__STRING_LENGTH]
    VAR_INPUT
        in : ULINT;
    END_VAR

    TO_STRING__ULINT := ULINT_TO_STRING(in);
END_FUNCTION

FUNCTION TO_STRING__BYTE : STRING[__STRING_LENGTH]
    VAR_INPUT
        in : BYTE;
    END_VAR

    TO_STRING__BYTE := BYTE_TO_STRING(in);
END_FUNCTION

FUNCTION TO_STRING__DWORD : STRING[__STRING_LENGTH]
    VAR_INPUT
        in : DWORD;
    END_VAR

    TO_STRING__DWORD := DWORD_TO_STRING(in);
END_FUNCTION

FUNCTION TO_STRING__LWORD : STRING[__STRING_LENGTH]
    VAR_INPUT
        in : LWORD;
    END_VAR

    TO_STRING__LWORD := LWORD_TO_STRING(in);
END_FUNCTION

FUNCTION TO_STRING__REAL : STRING[__STRING_LENGTH]
    VAR_INPUT
        in : REAL;
    END_VAR

    TO_STRING__REAL := REAL_TO_STRING(in);
END_FUNCTION

FUNCTION TO_STRING__LREAL : STRING[__STRING_LENGTH]
    VAR_INPUT
        in : LREAL;
    END_VAR

    TO_STRING__LREAL := LREAL_TO_STRING(in);
END_FUNCTION

FUNCTION TO_STRING__TIME : STRING[__STRING_LENGTH]
    VAR_INPUT
        in : TIME;
    END_VAR

    TO_STRING__TIME := TIME_TO_STRING(in);
END_FUNCTION

FUNCTION TO_STRING__LTIME : STRING[__STRING_LENGTH]
    VAR_INPUT
        in : LTIME;
    END_VAR

    TO_STRING__LTIME := LTIME_TO_STRING(in);
END_FUNCTION

FUNCTION TO_STRING__DATE : STRING[__STRING_LENGTH]
    VAR_INPUT
        in : DATE;
    END_VAR

    TO_STRING__DATE := DATE_TO_STRING(in);
END_FUNCTION

FUNCTION TO_STRING__LDATE : STRING[__STRING_LENGTH]
    VAR_INPUT
        in : LDATE;
    END_VAR

    TO_STRING__LDATE := LDATE_TO_STRING(in);
END_FUNCTION

FUNCTION TO_STRING__DT : STRING[__STRING_LENGTH]
    VAR_INPUT
        in : DT;
    END_VAR

    TO_STRING__DT := DT_TO_STRING(in);
END_FUNCTION

FUNCTION TO_STRING__LDT : STRING[__STRING_LENGTH]
    VAR_INPUT
        in : LDT;
    END_VAR

    TO_STRING__LDT := LDT_TO_STRING(in);
END_FUNCTION

FUNCTION TO_STRING__TOD : STRING[__STRING_LENGTH]
    VAR_INPUT
        in : TOD;
    END_VAR

    TO_STRING__TOD := TOD_TO_STRING(in);
END_FUNCTION

FUNCTION TO_STRING__LTOD : STRING[__STRING_LENGTH]
    VAR_INPUT
        in : LTOD;
    END_VAR

    TO_STRING__LTOD := LTOD_TO_STRING(in);
END_FUNCTION

// -----------------------------------------------------------------------------------------------------------
FUNCTION TO_WSTRING<T: ANY> : WSTRING[__STRING_LENGTH]
    VAR_INPUT
        in : T;
    END_VAR
END_FUNCTION

FUNCTION TO_WSTRING__WSTRING : WSTRING[__STRING_LENGTH]
    VAR_INPUT {ref}
        in : WSTRING;
    END_VAR

    TO_WSTRING__WSTRING := in;
END_FUNCTION

FUNCTION TO_WSTRING__STRING : WSTRING[__STRING_LENGTH]
    VAR_INPUT {ref}
        in : STRING;
    END_VAR

    STRING_TO_WSTRING_EXT(in, TO_WSTRING__STRING);
END_FUNCTION

FUNCTION TO_WSTRING__WCHAR : WSTRING[__STRING_LENGTH]
    VAR_INPUT
        in : WCHAR;
    END_VAR

    TO_WSTRING__WCHAR := WCHAR_TO_WSTRING(in);
END_FUNCTION

// Numeric, bit-string and date/time monomorphizations of the generic TO_WSTRING, each
// delegating to the corresponding typed <T>_TO_WSTRING conversion function.

FUNCTION TO_WSTRING__DINT : WSTRING[__STRING_LENGTH]
    VAR_INPUT
        in : DINT;
    END_VAR

    TO_WSTRING__DINT := DINT_TO_WSTRING(in);
END_FUNCTION

FUNCTION TO_WSTRING__LINT : WSTRING[__STRING_LENGTH]
    VAR_INPUT
        in : LINT;
    END_VAR

    TO_WSTRING__LINT := LINT_TO_WSTRING(in);
END_FUNCTION

FUNCTION TO_WSTRING__BYTE : WSTRING[__STRING_LENGTH]
    VAR_INPUT
        in : BYTE;
    END_VAR

    TO_WSTRING__BYTE := BYTE_TO_WSTRING(in);
END_FUNCTION

FUNCTION TO_WSTRING__DWORD : WSTRING[__STRING_LENGTH]
    VAR_INPUT
        in : DWORD;
    END_VAR

    TO_WSTRING__DWORD := DWORD_TO_WSTRING(in);
END_FUNCTION

FUNCTION TO_WSTRING__LWORD : WSTRING[__STRING_LENGTH]
    VAR_INPUT
        in : LWORD;
    END_VAR

    TO_WSTRING__LWORD := LWORD_TO_WSTRING(in);
END_FUNCTION

FUNCTION TO_WSTRING__REAL : WSTRING[__STRING_LENGTH]
    VAR_INPUT
        in : REAL;
    END_VAR

    TO_WSTRING__REAL := REAL_TO_WSTRING(in);
END_FUNCTION

FUNCTION TO_WSTRING__LREAL : WSTRING[__STRING_LENGTH]
    VAR_INPUT
        in : LREAL;
    END_VAR

    TO_WSTRING__LREAL := LREAL_TO_WSTRING(in);
END_FUNCTION

FUNCTION TO_WSTRING__TIME : WSTRING[__STRING_LENGTH]
    VAR_INPUT
        in : TIME;
    END_VAR

    TO_WSTRING__TIME := TIME_TO_WSTRING(in);
END_FUNCTION

FUNCTION TO_WSTRING__LTIME : WSTRING[__STRING_LENGTH]
    VAR_INPUT
        in : LTIME;
    END_VAR

    TO_WSTRING__LTIME := LTIME_TO_WSTRING(in);
END_FUNCTION

FUNCTION TO_WSTRING__DATE : WSTRING[__STRING_LENGTH]
    VAR_INPUT
        in : DATE;
    END_VAR

    TO_WSTRING__DATE := DATE_TO_WSTRING(in);
END_FUNCTION

FUNCTION TO_WSTRING__LDATE : WSTRING[__STRING_LENGTH]
    VAR_INPUT
        in : LDATE;
    END_VAR

    TO_WSTRING__LDATE := LDATE_TO_WSTRING(in);
END_FUNCTION

FUNCTION TO_WSTRING__DT : WSTRING[__STRING_LENGTH]
    VAR_INPUT
        in : DT;
    END_VAR

    TO_WSTRING__DT := DT_TO_WSTRING(in);
END_FUNCTION

FUNCTION TO_WSTRING__LDT : WSTRING[__STRING_LENGTH]
    VAR_INPUT
        in : LDT;
    END_VAR

    TO_WSTRING__LDT := LDT_TO_WSTRING(in);
END_FUNCTION

FUNCTION TO_WSTRING__TOD : WSTRING[__STRING_LENGTH]
    VAR_INPUT
        in : TOD;
    END_VAR

    TO_WSTRING__TOD := TOD_TO_WSTRING(in);
END_FUNCTION

FUNCTION TO_WSTRING__LTOD : WSTRING[__STRING_LENGTH]
    VAR_INPUT
        in : LTOD;
    END_VAR

    TO_WSTRING__LTOD := LTOD_TO_WSTRING(in);
END_FUNCTION

(* ---- to_string_conversions.st ---- *)
(******************************************************************************
*
* Converts native values to STRING and WSTRING.
*
******************************************************************************)
{external}
FUNCTION BOOL_TO_STRING : STRING[5]
VAR_INPUT
    IN : BOOL;
END_VAR
END_FUNCTION

FUNCTION BYTE_TO_STRING : STRING[3]
VAR_INPUT
    IN : BYTE;
END_VAR
    BYTE_TO_STRING_EXT(IN, BYTE_TO_STRING);
END_FUNCTION

{external}
FUNCTION BYTE_TO_STRING_EXT : DINT
VAR_INPUT
    IN : BYTE;
END_VAR
VAR_IN_OUT
    OUT : STRING[3];
END_VAR
END_FUNCTION

{external}
FUNCTION WORD_TO_STRING_EXT : DINT
VAR_INPUT
    IN : WORD;
END_VAR
VAR_IN_OUT
    OUT : STRING[5];
END_VAR
END_FUNCTION

FUNCTION WORD_TO_STRING : STRING[5]
VAR_INPUT
    IN : WORD;
END_VAR
    WORD_TO_STRING_EXT(IN, WORD_TO_STRING);
END_FUNCTION

{external}
FUNCTION LWORD_TO_STRING_EXT : DINT
VAR_INPUT
    IN : LWORD;
END_VAR
VAR_IN_OUT
    OUT : STRING[20];
END_VAR
END_FUNCTION

FUNCTION LWORD_TO_STRING : STRING[20]
VAR_INPUT
    IN : LWORD;
END_VAR
    LWORD_TO_STRING_EXT(IN, LWORD_TO_STRING);
END_FUNCTION

FUNCTION DWORD_TO_STRING : STRING[10]
VAR_INPUT
    IN : DWORD;
END_VAR
    DWORD_TO_STRING_EXT(IN, DWORD_TO_STRING);
END_FUNCTION

{external}
FUNCTION DWORD_TO_STRING_EXT : DINT
VAR_INPUT
    IN : DWORD;
END_VAR
VAR_IN_OUT
    OUT : STRING[10];
END_VAR
END_FUNCTION

{external}
FUNCTION LINT_TO_STRING_EXT : DINT
VAR_INPUT
    IN : LINT;
END_VAR
VAR_IN_OUT
    OUT : STRING[20];
END_VAR
END_FUNCTION

{external}
FUNCTION SINT_TO_STRING_EXT : DINT
VAR_INPUT
    IN : SINT;
END_VAR
VAR_IN_OUT
    OUT : STRING[4];
END_VAR
END_FUNCTION

FUNCTION SINT_TO_STRING : STRING[4]
VAR_INPUT
    IN : SINT;
END_VAR
    SINT_TO_STRING_EXT(IN, SINT_TO_STRING);
END_FUNCTION

{external}
FUNCTION INT_TO_STRING_EXT : DINT
VAR_INPUT
    IN : INT;
END_VAR
VAR_IN_OUT
    OUT : STRING[6];
END_VAR
END_FUNCTION

FUNCTION INT_TO_STRING : STRING[6]
VAR_INPUT
    IN : INT;
END_VAR
    INT_TO_STRING_EXT(IN, INT_TO_STRING);
END_FUNCTION

FUNCTION LINT_TO_STRING : STRING[20]
VAR_INPUT
    IN : LINT;
END_VAR
    LINT_TO_STRING_EXT(IN, LINT_TO_STRING);
END_FUNCTION

FUNCTION DINT_TO_STRING : STRING[11]
VAR_INPUT
    IN : DINT;
END_VAR
    DINT_TO_STRING_EXT(IN, DINT_TO_STRING);
END_FUNCTION

{external}
FUNCTION DINT_TO_STRING_EXT : DINT
VAR_INPUT
    IN : DINT;
END_VAR
VAR_IN_OUT
    OUT : STRING[11];
END_VAR
END_FUNCTION

FUNCTION USINT_TO_STRING : STRING[3]
VAR_INPUT
    IN : USINT;
END_VAR
    USINT_TO_STRING_EXT(IN, USINT_TO_STRING);
END_FUNCTION

{external}
FUNCTION USINT_TO_STRING_EXT : DINT
VAR_INPUT
    IN : USINT;
END_VAR
VAR_IN_OUT
    OUT : STRING[3];
END_VAR
END_FUNCTION

FUNCTION UINT_TO_STRING : STRING[5]
VAR_INPUT
    IN : UINT;
END_VAR
    UINT_TO_STRING_EXT(IN, UINT_TO_STRING);
END_FUNCTION

{external}
FUNCTION UINT_TO_STRING_EXT : DINT
VAR_INPUT
    IN : UINT;
END_VAR
VAR_IN_OUT
    OUT : STRING[5];
END_VAR
END_FUNCTION

FUNCTION UDINT_TO_STRING : STRING[10]
VAR_INPUT
    IN : UDINT;
END_VAR
    UDINT_TO_STRING_EXT(IN, UDINT_TO_STRING);
END_FUNCTION

{external}
FUNCTION UDINT_TO_STRING_EXT : DINT
VAR_INPUT
    IN : UDINT;
END_VAR
VAR_IN_OUT
    OUT : STRING[10];
END_VAR
END_FUNCTION

FUNCTION ULINT_TO_STRING : STRING[20]
VAR_INPUT
    IN : ULINT;
END_VAR
    ULINT_TO_STRING_EXT(IN, ULINT_TO_STRING);
END_FUNCTION

{external}
FUNCTION ULINT_TO_STRING_EXT : DINT
VAR_INPUT
    IN : ULINT;
END_VAR
VAR_IN_OUT
    OUT : STRING[20];
END_VAR
END_FUNCTION

{external}
FUNCTION LREAL_TO_STRING_EXT : DINT
VAR_INPUT
    IN : LREAL;
END_VAR
VAR_IN_OUT
    OUT : STRING[22];
END_VAR
END_FUNCTION

FUNCTION LREAL_TO_STRING : STRING[22]
VAR_INPUT
    IN : LREAL;
END_VAR
    LREAL_TO_STRING_EXT(IN, LREAL_TO_STRING);
END_FUNCTION

FUNCTION REAL_TO_STRING : STRING[22]
VAR_INPUT
    IN : REAL;
END_VAR
    LREAL_TO_STRING_EXT(IN, REAL_TO_STRING);
END_FUNCTION

{external}
FUNCTION DT_TO_STRING : STRING[22]
VAR_INPUT
    IN : DT;
END_VAR
END_FUNCTION

{external}
FUNCTION LDT_TO_STRING : STRING[33]
VAR_INPUT
    IN : LDT;
END_VAR
END_FUNCTION

{external}
FUNCTION TIME_TO_STRING : STRING[19]
VAR_INPUT
    IN : TIME;
END_VAR
END_FUNCTION

{external}
FUNCTION LTIME_TO_STRING : STRING[37]
VAR_INPUT
    IN : LTIME;
END_VAR
END_FUNCTION

{external}
FUNCTION DATE_TO_STRING : STRING[12]
VAR_INPUT
    IN : DATE;
END_VAR
END_FUNCTION

{external}
FUNCTION LDATE_TO_STRING : STRING[16]
VAR_INPUT
    IN : LDATE;
END_VAR
END_FUNCTION

{external}
FUNCTION TOD_TO_STRING : STRING[16]
VAR_INPUT
    IN : TOD;
END_VAR
END_FUNCTION

{external}
FUNCTION LTOD_TO_STRING : STRING[23]
VAR_INPUT
    IN : LTOD;
END_VAR
END_FUNCTION

FUNCTION DT_TO_WSTRING : WSTRING[__STRING_LENGTH]
VAR_INPUT
    IN : DT;
END_VAR
    STRING_TO_WSTRING_EXT(DT_TO_STRING(IN), DT_TO_WSTRING);
END_FUNCTION

FUNCTION LDT_TO_WSTRING : WSTRING[__STRING_LENGTH]
VAR_INPUT
    IN : LDT;
END_VAR
    STRING_TO_WSTRING_EXT(LDT_TO_STRING(IN), LDT_TO_WSTRING);
END_FUNCTION

FUNCTION TIME_TO_WSTRING : WSTRING[__STRING_LENGTH]
VAR_INPUT
    IN : TIME;
END_VAR
    STRING_TO_WSTRING_EXT(TIME_TO_STRING(IN), TIME_TO_WSTRING);
END_FUNCTION

FUNCTION LTIME_TO_WSTRING : WSTRING[__STRING_LENGTH]
VAR_INPUT
    IN : LTIME;
END_VAR
    STRING_TO_WSTRING_EXT(LTIME_TO_STRING(IN), LTIME_TO_WSTRING);
END_FUNCTION

FUNCTION DATE_TO_WSTRING : WSTRING[__STRING_LENGTH]
VAR_INPUT
    IN : DATE;
END_VAR
    STRING_TO_WSTRING_EXT(DATE_TO_STRING(IN), DATE_TO_WSTRING);
END_FUNCTION

FUNCTION LDATE_TO_WSTRING : WSTRING[__STRING_LENGTH]
VAR_INPUT
    IN : LDATE;
END_VAR
    STRING_TO_WSTRING_EXT(LDATE_TO_STRING(IN), LDATE_TO_WSTRING);
END_FUNCTION

FUNCTION TOD_TO_WSTRING : WSTRING[__STRING_LENGTH]
VAR_INPUT
    IN : TOD;
END_VAR
    STRING_TO_WSTRING_EXT(TOD_TO_STRING(IN), TOD_TO_WSTRING);
END_FUNCTION

FUNCTION LTOD_TO_WSTRING : WSTRING[__STRING_LENGTH]
VAR_INPUT
    IN : LTOD;
END_VAR
    STRING_TO_WSTRING_EXT(LTOD_TO_STRING(IN), LTOD_TO_WSTRING);
END_FUNCTION

FUNCTION BYTE_TO_WSTRING : WSTRING[__STRING_LENGTH]
VAR_INPUT
    IN : BYTE;
END_VAR
    STRING_TO_WSTRING_EXT(BYTE_TO_STRING(IN), BYTE_TO_WSTRING);
END_FUNCTION

FUNCTION LWORD_TO_WSTRING : WSTRING[__STRING_LENGTH]
VAR_INPUT
    IN : LWORD;
END_VAR
    STRING_TO_WSTRING_EXT(LWORD_TO_STRING(IN), LWORD_TO_WSTRING);
END_FUNCTION

FUNCTION DWORD_TO_WSTRING : WSTRING[__STRING_LENGTH]
VAR_INPUT
    IN : DWORD;
END_VAR
    DWORD_TO_WSTRING := LWORD_TO_WSTRING(IN);
END_FUNCTION

FUNCTION LINT_TO_WSTRING : WSTRING[__STRING_LENGTH]
VAR_INPUT
    IN : LINT;
END_VAR
    STRING_TO_WSTRING_EXT(LINT_TO_STRING(IN), LINT_TO_WSTRING);
END_FUNCTION

FUNCTION DINT_TO_WSTRING : WSTRING[__STRING_LENGTH]
VAR_INPUT
    IN : DINT;
END_VAR
    DINT_TO_WSTRING := LINT_TO_WSTRING(IN);
END_FUNCTION

FUNCTION LREAL_TO_WSTRING : WSTRING[__STRING_LENGTH]
VAR_INPUT
    IN : LREAL;
END_VAR
    STRING_TO_WSTRING_EXT(LREAL_TO_STRING(IN), LREAL_TO_WSTRING);
END_FUNCTION

FUNCTION REAL_TO_WSTRING : WSTRING[__STRING_LENGTH]
VAR_INPUT
    IN : REAL;
END_VAR
    REAL_TO_WSTRING := LREAL_TO_WSTRING(IN);
END_FUNCTION

(* ---- trunc_int.st ---- *)
(********************
*
* Converts a floating point number to SINT
*
********************)
FUNCTION TRUNC_SINT<T: ANY_REAL> : SINT
    VAR_INPUT
        in : T;
    END_VAR
END_FUNCTION

(********************
*
* Converts REAL to SINT
*
********************)
FUNCTION TRUNC_SINT__REAL : SINT
    VAR_INPUT
        in : REAL;
    END_VAR

    TRUNC_SINT__REAL := in;
END_FUNCTION

(********************
*
* Converts LREAL to SINT
*
********************)
FUNCTION TRUNC_SINT__LREAL : SINT
    VAR_INPUT
        in : LREAL;
    END_VAR

    TRUNC_SINT__LREAL := in;
END_FUNCTION

(********************
*
* Converts a floating point number to USINT
*
********************)
FUNCTION TRUNC_USINT<T: ANY_REAL> : USINT
    VAR_INPUT
        in : T;
    END_VAR
END_FUNCTION

(********************
*
* Converts REAL to USINT
*
********************)
FUNCTION TRUNC_USINT__REAL : USINT
    VAR_INPUT
        in : REAL;
    END_VAR

    TRUNC_USINT__REAL := in;
END_FUNCTION

(********************
*
* Converts LREAL to USINT
*
********************)
FUNCTION TRUNC_USINT__LREAL : USINT
    VAR_INPUT
        in : LREAL;
    END_VAR

    TRUNC_USINT__LREAL := in;
END_FUNCTION

(********************
*
* Converts a floating point number to INT
*
********************)
FUNCTION TRUNC_INT<T: ANY_REAL> : INT
    VAR_INPUT
        in : T;
    END_VAR
END_FUNCTION

(********************
*
* Converts REAL to INT
*
********************)
FUNCTION TRUNC_INT__REAL : INT
    VAR_INPUT
        in : REAL;
    END_VAR

    TRUNC_INT__REAL := in;
END_FUNCTION

(********************
*
* Converts LREAL to INT
*
********************)
FUNCTION TRUNC_INT__LREAL : INT
    VAR_INPUT
        in : LREAL;
    END_VAR

    TRUNC_INT__LREAL := in;
END_FUNCTION

(********************
*
* Converts a floating point number to UINT
*
********************)
FUNCTION TRUNC_UINT<T: ANY_REAL> : UINT
    VAR_INPUT
        in : T;
    END_VAR
END_FUNCTION

(********************
*
* Converts REAL to UINT
*
********************)
FUNCTION TRUNC_UINT__REAL : UINT
    VAR_INPUT
        in : REAL;
    END_VAR

    TRUNC_UINT__REAL := in;
END_FUNCTION

(********************
*
* Converts LREAL to UINT
*
********************)
FUNCTION TRUNC_UINT__LREAL : UINT
    VAR_INPUT
        in : LREAL;
    END_VAR

    TRUNC_UINT__LREAL := in;
END_FUNCTION

(********************
*
* Converts a floating point number to DINT
*
********************)
FUNCTION TRUNC_DINT<T: ANY_REAL> : DINT
    VAR_INPUT
        in : T;
    END_VAR
END_FUNCTION

(********************
*
* Converts REAL to DINT
*
********************)
FUNCTION TRUNC_DINT__REAL : DINT
    VAR_INPUT
        in : REAL;
    END_VAR

    TRUNC_DINT__REAL := in;
END_FUNCTION

(********************
*
* Converts LREAL to DINT
*
********************)
FUNCTION TRUNC_DINT__LREAL : DINT
    VAR_INPUT
        in : LREAL;
    END_VAR

    TRUNC_DINT__LREAL := in;
END_FUNCTION

(********************
*
* Converts a floating point number to UDINT
*
********************)
FUNCTION TRUNC_UDINT<T: ANY_REAL> : UDINT
    VAR_INPUT
        in : T;
    END_VAR
END_FUNCTION

(********************
*
* Converts REAL to UDINT
*
********************)
FUNCTION TRUNC_UDINT__REAL : UDINT
    VAR_INPUT
        in : REAL;
    END_VAR

    TRUNC_UDINT__REAL := in;
END_FUNCTION

(********************
*
* Converts LREAL to UDINT
*
********************)
FUNCTION TRUNC_UDINT__LREAL : UDINT
    VAR_INPUT
        in : LREAL;
    END_VAR

    TRUNC_UDINT__LREAL := in;
END_FUNCTION

(********************
*
* Converts a floating point number to LINT
*
********************)
FUNCTION TRUNC_LINT<T: ANY_REAL> : LINT
    VAR_INPUT
        in : T;
    END_VAR
END_FUNCTION

(********************
*
* Converts REAL to LINT
*
********************)
FUNCTION TRUNC_LINT__REAL : LINT
    VAR_INPUT
        in : REAL;
    END_VAR

    TRUNC_LINT__REAL := in;
END_FUNCTION

(********************
*
* Converts LREAL to LINT
*
********************)
FUNCTION TRUNC_LINT__LREAL : LINT
    VAR_INPUT
        in : LREAL;
    END_VAR

    TRUNC_LINT__LREAL := in;
END_FUNCTION

(********************
*
* Converts a floating point number to ULINT
*
********************)
FUNCTION TRUNC_ULINT<T: ANY_REAL> : ULINT
    VAR_INPUT
        in : T;
    END_VAR
END_FUNCTION

(********************
*
* Converts REAL to ULINT
*
********************)
FUNCTION TRUNC_ULINT__REAL : ULINT
    VAR_INPUT
        in : REAL;
    END_VAR

    TRUNC_ULINT__REAL := in;
END_FUNCTION

(********************
*
* Converts LREAL to ULINT
*
********************)
FUNCTION TRUNC_ULINT__LREAL : ULINT
    VAR_INPUT
        in : LREAL;
    END_VAR

    TRUNC_ULINT__LREAL := in;
END_FUNCTION

(* ---- validation_functions.st ---- *)
(******************************************************************************
Description: Validation function for ANY_REAL
Input:
  - IN: ANY_REAL
Return:
  - FALSE: If input is Not-a-Number(NaN) or infinite(+Inf, -Inf)
  - TRUE: Otherwise
******************************************************************************)
{external}
FUNCTION IS_VALID <T: ANY_REAL> : BOOL
VAR_INPUT
    IN : T;
END_VAR
END_FUNCTION

(******************************************************************************
Description: Validation function for ANY_BIT
Validate if the binary representation of the input
would result in a valid BCD representation
Input:
  - IN: ANY_BIT
Return:
  - TRUE: The value of each 4bits represented digit must be between 0-9
  - FALSE: If the value of any 4bits represented digit is higher than 9
******************************************************************************)
{external}
FUNCTION IS_VALID_BCD <T: ANY_BIT> : BOOL
VAR_INPUT
    IN : T;
END_VAR
END_FUNCTION

(* ---- bistable_functionblocks.st ---- *)
(******************************************************************************
Description: Bistable function, set dominant
Input:
  - SET1: Dominant input of bistable function
  - RESET: Input of bistable function
Output:
  - Q1: Result of bistable function
Return: Output is used as return
******************************************************************************)
{external}
FUNCTION_BLOCK SR
VAR_INPUT
    SET1: BOOL;
    RESET: BOOL;
END_VAR
VAR_OUTPUT
    Q1: BOOL;
END_VAR
END_FUNCTION_BLOCK

(******************************************************************************
Description: Bistable function, reset dominant
Input:
  - SET: Input of bistable function
  - RESET1: Dominant input of bistable function
Output:
  - Q1: Result of bistable function
Return: Output is used as return
******************************************************************************)
{external}
FUNCTION_BLOCK RS
VAR_INPUT
    SET:    BOOL;
    RESET1: BOOL;
END_VAR
VAR_OUTPUT
    Q1:     BOOL;
END_VAR
END_FUNCTION_BLOCK
